      $ 2072 "Vial_liq_pick_3" "breakAfter"
      movel(Vial_liq_pick_3_p, a=0.5, v=0.1)
      $ 2073 "Vial_liq_pick_4" "breakAfter"
      movel(Vial_liq_pick_4_p, a=0.5, v=0.1)
      # begin: URCap Program Node
      #   Source: Robotiq_Grippers, 3.17.0.105337, Robotiq Inc.
      #   Type: Gripper
      $ 2074 "Gripper Close (1)"
      if not(gripper_connected[0]):
        popup("Gripper 1 must be connected to run this program.", "No connection", False, True, True)
      end
      if not(rq_is_gripper_activated("1")):
        popup("Gripper 1 is not activated. Go to Installation tab > Gripper to activate it and run the program again.", "Not activated", False, True, True)
      end
      rq_set_pos_spd_for(255, 82, 71, "1")
      rq_wait_pos_spe_for_request(255, 82, 71, "1")
      rq_go_to("1")
      rq_wait("1")
      # end: URCap Program Node
      $ 2075 "Wait: 1.0"
      sleep(1.0)
      $ 2076 "Set GRP_3F_Open=On"
      set_standard_digital_out(5, True)
      $ 2077 "Wait: 0.5"
      sleep(0.5)
      $ 2078 "Vial_liq_abov_2" "breakAfter"
      movel(Vial_liq_abov_2_p, a=0.3, v=0.05, r=0.05)
      $ 2079 "MoveL"
      $ 2080 "Liquid_midway_1" "breakAfter"
      movel(Liquid_midway_1_p, a=0.5, v=0.1)
      $ 2081 "Loop 3 times"
      Loop_1 = 0
      while (Loop_1 < 3):
        $ 2082 "shake_3" "breakAfter"
        movel(shake_3_p, a=2.0, v=0.5)
        $ 2083 "shake_4" "breakAfter"
        movel(shake_4_p, a=2.0, v=0.5)
        Loop_1 = Loop_1 + 1
      end
      $ 2084 "drop_above_3" "breakAfter"
      movel(drop_above_3_p, a=0.5, v=0.1)
      $ 2085 "drop_above_4" "breakAfter"
      movel(drop_above_4_p, a=0.5, v=0.1)
      $ 2086 "liq_tran_3" "breakAfter"
      movel(liq_tran_3_p, a=0.5, v=0.05, r=0.008)
      $ 2087 "Wait: 1.0"
      sleep(1.0)
      $ 2088 "drop_above_5" "breakAfter"
      movel(drop_above_5_p, a=0.5, v=0.1)
      $ 2089 "Waypoint_92" "breakAfter"
      movel(Waypoint_92_p, a=0.5, v=0.1)
      $ 2090 "liq_tran_4" "breakAfter"
      movel(liq_tran_4_p, a=0.5, v=0.05)
      $ 2091 "Wait: 1.0"
      sleep(1.0)
      $ 2092 "drop_above_6" "breakAfter"
      movel(drop_above_6_p, a=0.5, v=0.1)
      $ 2093 "drop_above_7" "breakAfter"
      movel(drop_above_7_p, a=0.5, v=0.1)
      $ 2094 "Liquid_midway_2" "breakAfter"
      movel(Liquid_midway_2_p, a=0.5, v=0.1)
      $ 2095 "MoveL"
      $ 2096 "Vial_drop_abo_1" "breakAfter"
      movel(Vial_drop_abo_1_p, a=0.5, v=0.1)
      $ 2097 "Vial_liq_drop_1" "breakAfter"
      movel(Vial_liq_drop_1_p, a=0.5, v=0.1)
      # begin: URCap Program Node
      #   Source: Robotiq_Grippers, 3.17.0.105337, Robotiq Inc.
      #   Type: Gripper
      $ 2098 "Gripper Open (1)"
      if not(gripper_connected[0]):
        popup("Gripper 1 must be connected to run this program.", "No connection", False, True, True)
      end
      if not(rq_is_gripper_activated("1")):
        popup("Gripper 1 is not activated. Go to Installation tab > Gripper to activate it and run the program again.", "Not activated", False, True, True)
      end
      rq_set_pos_spd_for(0, 82, 71, "1")
      rq_wait_pos_spe_for_request(0, 82, 71, "1")
      rq_go_to("1")
      rq_wait("1")
      # end: URCap Program Node
      $ 2099 "Vial_drop_abo_2" "breakAfter"
      movel(Vial_drop_abo_2_p, a=0.5, v=0.1)
    elif (34 == switch_1):
      $ 2100 "Case 34"
      $ 2101 "Task≔'Dosing'"
      global Task="Dosing"
      $ 2102 "tilt_to_home()"
      tilt_to_home()
      $ 2103 "Powder dosing all"
      $ 2104 "tilt_angle_sent≔0.0"
      global tilt_angle_sent=0.0
      $ 2105 "send_target_info()"
      send_target_info()
      $ 2107 "prev_spat≔''"
      global prev_spat=""
      $ 2108 "spatula≔''"
      global spatula=""
      $ 2109 "scoop_status≔'normal'"
      global scoop_status="normal"
      $ 2110 "send_powder_info()"
      send_powder_info()
      $ 2111 "Set AO[0]=0.0"
      set_standard_analog_out(0, 0.0)
      $ 2112 "Wait: 0.2"
      sleep(0.2)
      $ 2113 "reach pots decapping pose"
      # begin: URCap Program Node
      #   Source: SensoPart VISOR Robotic, 2.0.6, SensoPart Industriesensorik GmbH
      #   Type: VISOR Robotic App
      $ 2119 "VISOR Easy Pick"
      def visorFuncEasyPick_5caf8b():
        # begin: URCap Program Node
        #   Source: SensoPart VISOR Robotic, 2.0.6, SensoPart Industriesensorik GmbH
        #   Type: Easy Pick Setup
        $ 2120 "# 1 Setup" "noBreak"
        local easyPickVisorId = 1
        local easyPickArmMounted = True
        local easyPickSetJob = True
        local easyPickJobName = "Weight_scale"
        local easyPickAtImgAcq = False
        local easyPickImgAcqPose = Trigger
        # end: URCap Program Node
        # begin: URCap Program Node
        #   Source: SensoPart VISOR Robotic, 2.0.6, SensoPart Industriesensorik GmbH
        #   Type: Process
        $ 2121 "Process" "noBreak"
        local easyPickObjTaken = False
        local easyPickTrigger = False
        local easyPickPoseIdx = 0
        local easyPickPose = p[0,0,0,0,0,0]
        def easyPickFuncTrigger(visorId, setJob, jobName, arm):
        if (setJob):
          visor_changeJob(visorId, jobName, 6000)
        end
        if (arm):
          visor_trigger(visorId, 6000, "arm")
        else:
          visor_trigger(visorId, 6000)
        end
        global easyPickParts_4=visor_partsFound(visorId)
        visor_easyPickUpdate(visorId, "parts", visor_partsFound(visorId))
        return visor_getPose3d(visorId, 0)
      end
      while (not easyPickObjTaken):
        easyPickTrigger = (easyPickCount_4 >= visor_partsFound(easyPickVisorId)) or (easyPickCount_4 > 9) or (not visor_easyPickCheckIdent("a98771", easyPickVisorId))
        if (easyPickTrigger):
          easyPickCount_4 = 0
        end
        easyPickPoseIdx = easyPickCount_4
        easyPickPose = visor_getPose3d(easyPickVisorId, easyPickPoseIdx)
        visor_easyPickUpdate(easyPickVisorId, "counter", easyPickPoseIdx)
        # begin: URCap Program Node
        #   Source: SensoPart VISOR Robotic, 2.0.6, SensoPart Industriesensorik GmbH
        #   Type: Image Acquisition Pose
        $ 2122 "Image Acquisition Pose" "noBreak"
        if (easyPickTrigger):
          if (not easyPickAtImgAcq):
            movej(pose_trans(easyPickImgAcqPose,p[0.0000,0.0000,-0.0000,0.0000,0.0000,0.0000]),a=1.3963,v=1.0472,t=0.000000,r=0.000000)
            easyPickAtImgAcq = True
          end
          easyPickPose = easyPickFuncTrigger(easyPickVisorId, easyPickSetJob, easyPickJobName, easyPickArmMounted)
        end
        # end: URCap Program Node
        # begin: URCap Program Node
        #   Source: SensoPart VISOR Robotic, 2.0.6, SensoPart Industriesensorik GmbH
        #   Type: Object Detected
        $ 2123 "Object Detected" "noBreak"
        if (visor_partsFound(easyPickVisorId) > 0):
          $ 2124 "Open Gripper" "noBreak"
          $ 2125 "weight_value≔get_weight()" "noBreak"
          global weight_value=get_weight()
          $ 2126 "Wait: 0.5" "noBreak"
          sleep(0.5)
          $ 2127 "diff≔target_weight-weight_value" "noBreak"
          global diff=target_weight-weight_value
          $ 2128 "compute_level_percent(W_now, weight_value)" "noBreak"
          compute_level_percent(W_now, weight_value)
          $ 2129 "send_level_info()" "noBreak"
          send_level_info()
          $ 2130 "spatula≔select_spatula(Flowability, level, diff, bulk_density, mouth_d)" "noBreak"
          global spatula=select_spatula(Flowability, level, diff, bulk_density, mouth_d)
          $ 2131 "Wait: 0.2" "noBreak"
          sleep(0.2)
          $ 2132 "send_spatula_info()" "noBreak"
          send_spatula_info()
          $ 2133 "Pick spatula" "noBreak"
          $ 2134 "If spatula ≟ 'spatula_L'" "noBreak"
          if (spatula  ==  "spatula_L"):
            $ 2135 "MoveJ" "noBreak"
            $ 2136 "Spatula_otw" "noBreak"
            movej(get_inverse_kin(Spatula_otw_p, qnear=Spatula_otw_q), a=1.3962634015954636, v=1.0471975511965976)
            $ 2137 "pick_spat_L_abv" "noBreak"
            movej(get_inverse_kin(pick_spat_L_abv_p, qnear=pick_spat_L_abv_q), a=1.3962634015954636, v=1.0471975511965976)
            $ 2138 "MoveL" "noBreak"
            $ 2139 "spat_L_pick" "noBreak"
            movel(spat_L_pick_p, a=1.2, v=0.25)
            # begin: URCap Program Node
            #   Source: Robotiq_Grippers, 3.17.0.105337, Robotiq Inc.
            #   Type: Gripper
            $ 2140 "Gripper Close (1)" "noBreak"
            if not(gripper_connected[0]):
              popup("Gripper 1 must be connected to run this program.", "No connection", False, True, True)
            end
            if not(rq_is_gripper_activated("1")):
              popup("Gripper 1 is not activated. Go to Installation tab > Gripper to activate it and run the program again.", "Not activated", False, True, True)
            end
            rq_set_pos_spd_for(255, 0, 77, "1")
            rq_wait_pos_spe_for_request(255, 0, 77, "1")
            rq_go_to("1")
            rq_wait("1")
            # end: URCap Program Node
            $ 2141 "spat_L_lift" "noBreak"
            movel(spat_L_lift_p, a=1.2, v=0.25, r=0.01)
            $ 2142 "spat_L_side" "noBreak"
            movel(spat_L_side_p, a=1.2, v=0.25, r=0.01)
            $ 2143 "spat_L_up" "noBreak"
            movel(spat_L_up_p, a=1.2, v=0.25, r=0.05)
            $ 2144 "MoveJ" "noBreak"
            $ 2145 "Spatula_otw" "noBreak"
            movej(get_inverse_kin(Spatula_otw_p, qnear=Spatula_otw_q), a=1.3962634015954636, v=1.0471975511965976)
          else:
            $ 2146 "ElseIf spatula ≟'spatula_M'" "noBreak"
            if (spatula  == "spatula_M"):
              $ 2147 "MoveJ" "noBreak"
              $ 2148 "Spatula_otw" "noBreak"
              movej(get_inverse_kin(Spatula_otw_p, qnear=Spatula_otw_q), a=1.3962634015954636, v=1.0471975511965976)
              $ 2149 "spat_M_up" "noBreak"
              movej(get_inverse_kin(spat_M_up_p, qnear=spat_M_up_q), a=1.3962634015954636, v=1.0471975511965976, r=0.05)
              $ 2150 "MoveL" "noBreak"
              $ 2151 "spat_M_pick" "noBreak"
              movel(spat_M_pick_p, a=1.2, v=0.25)
              # begin: URCap Program Node
              #   Source: Robotiq_Grippers, 3.17.0.105337, Robotiq Inc.
              #   Type: Gripper
              $ 2152 "Gripper Close (1)" "noBreak"
              if not(gripper_connected[0]):
                popup("Gripper 1 must be connected to run this program.", "No connection", False, True, True)
              end
              if not(rq_is_gripper_activated("1")):
                popup("Gripper 1 is not activated. Go to Installation tab > Gripper to activate it and run the program again.", "Not activated", False, True, True)
              end
              rq_set_pos_spd_for(255, 0, 77, "1")
              rq_wait_pos_spe_for_request(255, 0, 77, "1")
              rq_go_to("1")
              rq_wait("1")
              # end: URCap Program Node
              $ 2153 "spat_M_up" "noBreak"
              movel(spat_M_up_p, a=1.2, v=0.25, r=0.05)
              $ 2154 "Spatula_otw" "noBreak"
              movel(Spatula_otw_p, a=1.2, v=0.25)
              $ 2155 "switch_spat_M≔ False " "noBreak"
              global switch_spat_M=  False
            else:
              $ 2156 "ElseIf spatula≟'spatula_S'" "noBreak"
              if (spatula == "spatula_S"):
                $ 2157 "MoveJ" "noBreak"
                $ 2158 "Spatula_otw" "noBreak"
                movej(get_inverse_kin(Spatula_otw_p, qnear=Spatula_otw_q), a=1.3962634015954636, v=1.0471975511965976)
                $ 2159 "spat_S_Up_7" "noBreak"
                movej(get_inverse_kin(spat_S_Up_7_p, qnear=spat_S_Up_7_q), a=1.3962634015954636, v=1.0471975511965976, r=0.05)
                $ 2160 "MoveL" "noBreak"
                $ 2161 "spat_S_Pick_4" "noBreak"
                movel(spat_S_Pick_4_p, a=1.2, v=0.25)
                # begin: URCap Program Node
                #   Source: Robotiq_Grippers, 3.17.0.105337, Robotiq Inc.
                #   Type: Gripper
                $ 2162 "Gripper Close (1)" "noBreak"
                if not(gripper_connected[0]):
                  popup("Gripper 1 must be connected to run this program.", "No connection", False, True, True)
                end
                if not(rq_is_gripper_activated("1")):
                  popup("Gripper 1 is not activated. Go to Installation tab > Gripper to activate it and run the program again.", "Not activated", False, True, True)
                end
                rq_set_pos_spd_for(255, 0, 77, "1")
                rq_wait_pos_spe_for_request(255, 0, 77, "1")
                rq_go_to("1")
                rq_wait("1")
                # end: URCap Program Node
                $ 2163 "spat_S_Up_8" "noBreak"
                movel(spat_S_Up_8_p, a=1.2, v=0.25, r=0.05)
                $ 2164 "Spatula_otw" "noBreak"
                movel(Spatula_otw_p, a=1.2, v=0.25)
                $ 2165 "switch_spat_S≔ False " "noBreak"
                global switch_spat_S=  False
              else:
                $ 2166 "ElseIf spatula≟'spatula_flat_M'" "noBreak"
                if (spatula == "spatula_flat_M"):
                  $ 2167 "MoveJ" "noBreak"
                  $ 2168 "Spatula_otw" "noBreak"
                  movej(get_inverse_kin(Spatula_otw_p, qnear=Spatula_otw_q), a=1.3962634015954636, v=1.0471975511965976)
                  $ 2169 "spat_flatM_up" "noBreak"
                  movej(get_inverse_kin(spat_flatM_up_p, qnear=spat_flatM_up_q), a=1.3962634015954636, v=1.0471975511965976, r=0.05)
                  $ 2170 "MoveL" "noBreak"
                  $ 2171 "spat_flatM_pick" "noBreak"
                  movel(spat_flatM_pick_p, a=1.2, v=0.25)
                  # begin: URCap Program Node
                  #   Source: Robotiq_Grippers, 3.17.0.105337, Robotiq Inc.
                  #   Type: Gripper
                  $ 2172 "Gripper Close (1)" "noBreak"
                  if not(gripper_connected[0]):
                    popup("Gripper 1 must be connected to run this program.", "No connection", False, True, True)
                  end
                  if not(rq_is_gripper_activated("1")):
                    popup("Gripper 1 is not activated. Go to Installation tab > Gripper to activate it and run the program again.", "Not activated", False, True, True)
                  end
                  rq_set_pos_spd_for(255, 0, 77, "1")
                  rq_wait_pos_spe_for_request(255, 0, 77, "1")
                  rq_go_to("1")
                  rq_wait("1")
                  # end: URCap Program Node
                  $ 2173 "spat_flatM_up" "noBreak"
                  movel(spat_flatM_up_p, a=1.2, v=0.25, r=0.05)
                  $ 2174 "Spatula_otw" "noBreak"
                  movel(Spatula_otw_p, a=1.2, v=0.25)
                  $ 2175 "switch_spat_F_M≔ False " "noBreak"
                  global switch_spat_F_M=  False
                else:
                  $ 2176 "ElseIf spatula≟'spatula_flat_S'" "noBreak"
                  if (spatula == "spatula_flat_S"):
                    $ 2177 "MoveJ" "noBreak"
                    $ 2178 "Spatula_otw" "noBreak"
                    movej(get_inverse_kin(Spatula_otw_p, qnear=Spatula_otw_q), a=1.3962634015954636, v=1.0471975511965976)
                    $ 2179 "spat_flatS_up" "noBreak"
                    movej(get_inverse_kin(spat_flatS_up_p, qnear=spat_flatS_up_q), a=1.3962634015954636, v=1.0471975511965976, r=0.05)
                    $ 2180 "MoveL" "noBreak"
                    $ 2181 "spat_flatS_pick" "noBreak"
                    movel(spat_flatS_pick_p, a=1.2, v=0.25)
                    # begin: URCap Program Node
                    #   Source: Robotiq_Grippers, 3.17.0.105337, Robotiq Inc.
                    #   Type: Gripper
                    $ 2182 "Gripper Close (1)" "noBreak"
                    if not(gripper_connected[0]):
                      popup("Gripper 1 must be connected to run this program.", "No connection", False, True, True)
                    end
                    if not(rq_is_gripper_activated("1")):
                      popup("Gripper 1 is not activated. Go to Installation tab > Gripper to activate it and run the program again.", "Not activated", False, True, True)
                    end
                    rq_set_pos_spd_for(255, 0, 77, "1")
                    rq_wait_pos_spe_for_request(255, 0, 77, "1")
                    rq_go_to("1")
                    rq_wait("1")
                    # end: URCap Program Node
                    $ 2183 "spat_flatS_up" "noBreak"
                    movel(spat_flatS_up_p, a=1.2, v=0.25, r=0.05)
                    $ 2184 "Spatula_otw" "noBreak"
                    movel(Spatula_otw_p, a=1.2, v=0.25)
                    $ 2185 "switch_spat_F_S≔ False " "noBreak"
                    global switch_spat_F_S=  False
                  end
                end
              end
            end
          end
          $ 2186 "Action_Info≔'Scooping'" "noBreak"
          global Action_Info="Scooping"
          $ 2187 "auto_tilt_and_scoop(W_now, target_weight, weight_value)" "noBreak"
          auto_tilt_and_scoop(W_now, target_weight, weight_value)
          $ 2188 "Action_Info≔'Dosing'" "noBreak"
          global Action_Info="Dosing"
          # begin: URCap Program Node
          #   Source: SensoPart VISOR Robotic, 2.0.6, SensoPart Industriesensorik GmbH
          #   Type: Approach Pose
          $ 2189 "Approach Pose" "noBreak"
          movej(pose_trans(easyPickPose,p[0.0000,0.0000,-0.0000,0.0000,0.0000,0.0000]),a=0.2618,v=0.1745,t=0.000000,r=0.000000)
          # end: URCap Program Node
          # begin: URCap Program Node
          #   Source: SensoPart VISOR Robotic, 2.0.6, SensoPart Industriesensorik GmbH
          #   Type: Target Pose
          $ 2190 "Target Pose" "noBreak"
          movel(pose_trans(easyPickPose,p[0.0000,0.0000,-0.0000,0.0000,0.0000,0.0000]),a=0.0500,v=0.0200,t=0.000000,r=0.000000)
          # end: URCap Program Node
          $ 2191 "Close Gripper" "noBreak"
          $ 2192 "current_p≔get_actual_tcp_pose()" "noBreak"
          global current_p= get_actual_tcp_pose ()
          $ 2193 "dispense_pos≔pose_trans(current_p,p[0,0,0,0,-deg2rad(spatula_ry),0])" "noBreak"
          global dispense_pos=pose_trans(current_p,p[0,0,0,0,-deg2rad(spatula_ry),0])
          $ 2195 "Loop weight_value≤target_weight " "noBreak"
          thread Thread_while_2195():
            while (True):
              $ 2196 "MoveL" "noBreak"
              $ 2197 "dispense_pos" "noBreak"
              movel(dispense_pos, a=0.2, v=0.1)
              $ 2198 "log_weight()" "noBreak"
              log_weight()
              $ 2200 "CCW_full_Rotate()" "noBreak"
              CCW_full_Rotate()
              $ 2201 "Start_thread≔ True " "noBreak"
              global Start_thread=  True
              $ 2202 "vib_thread≔ True " "noBreak"
              global vib_thread=  True
              $ 2203 "Wait: 0.5" "noBreak"
              sleep(0.5)
              $ 2204 "If diff ≥(target_g*1.2)" "noBreak"
              if (diff  >= (target_g*1.2)):
                $ 2205 "tilt_pose≔pose_trans(get_actual_tcp_pose(), p[0, 0, 0, 0, 0, 2.0])" "noBreak"
                global tilt_pose=pose_trans(get_actual_tcp_pose(), p[0, 0, 0, 0, 0, 2.0])
                $ 2206 "movel(tilt_pose, a=0.5, v=0.5, r=0.00001)" "noBreak"
                movel(tilt_pose, a=0.5, v=0.5, r=0.00001)
              else:
                $ 2207 "Else" "noBreak"
                $ 2208 "Loop weight_value≤(target_weight-0.00) and tilt_angle≥(-1.999) and tilt_angle≤0.5" "noBreak"
                thread Thread_while_2208():
                  while (True):
                    $ 2209 "current_error≔target_weight-weight_value" "noBreak"
                    global current_error=target_weight-weight_value
                    $ 2210 "Integral_error≔Integral_error+current_error*dt" "noBreak"
                    global Integral_error=Integral_error+current_error*dt
                    $ 2211 "derivative≔(current_error-previous_error)/dt" "noBreak"
                    global derivative=(current_error-previous_error)/dt
                    $ 2212 "tilt_increment≔(kp*current_error)+(ki*Integral_error)+(kd*derivative)" "noBreak"
                    global tilt_increment=(kp*current_error)+(ki*Integral_error)+(kd*derivative)
                    $ 2213 "current_pose≔get_actual_tcp_pose()" "noBreak"
                    global current_pose= get_actual_tcp_pose ()
                    $ 2214 "tilt_angle≔current_pose[5]" "noBreak"
                    global tilt_angle=current_pose[5]
                    $ 2215 "tilt_pose≔pose_trans(current_pose, p[0, 0, 0, 0, 0, tilt_increment])" "noBreak"
                    global tilt_pose=pose_trans(current_pose, p[0, 0, 0, 0, 0, tilt_increment])
                    $ 2216 "movel(tilt_pose, a=0.1, v=0.1, r=0.00001)" "noBreak"
                    movel(tilt_pose, a=0.1, v=0.1, r=0.00001)
                    $ 2217 "previous_error≔current_error" "noBreak"
                    global previous_error=current_error
                  end
                end
                if (weight_value <= (target_weight-0.00)  and  tilt_angle >= (-1.999)  and  tilt_angle <= 0.5):
                  global thread_handler_2208=run Thread_while_2208()
                  while (weight_value <= (target_weight-0.00)  and  tilt_angle >= (-1.999)  and  tilt_angle <= 0.5):
                    sync()
                  end
                  kill thread_handler_2208
                end
              end
              $ 2218 "weight_value≔get_weight()" "noBreak"
              global weight_value=get_weight()
              $ 2220 "tilt_angle≔-1" "noBreak"
              global tilt_angle=-1
              $ 2221 "Wait: 0.5" "noBreak"
              sleep(0.5)
              $ 2222 "Start_thread≔ False " "noBreak"
              global Start_thread=  False
              $ 2223 "vib_thread≔ False " "noBreak"
              global vib_thread=  False
              $ 2225 "dispense_pos" "noBreak"
              movel(dispense_pos, a=1.2, v=0.25)
              $ 2226 "compute_level_percent(W_now, weight_value)" "noBreak"
              compute_level_percent(W_now, weight_value)
              $ 2227 "prev_spat≔spatula" "noBreak"
              global prev_spat=spatula
              $ 2228 "Wait: 0.2" "noBreak"
              sleep(0.2)
              $ 2229 "spatula≔select_spatula(Flowability, level, diff, bulk_density, mouth_d)" "noBreak"
              global spatula=select_spatula(Flowability, level, diff, bulk_density, mouth_d)
              $ 2230 "Wait: 1.0" "noBreak"
              sleep(1.0)
              $ 2231 "send_level_info()" "noBreak"
              send_level_info()
              $ 2232 "send_spatula_info()" "noBreak"
              send_spatula_info()
              $ 2233 "Integral_error≔0" "noBreak"
              global Integral_error=0
              $ 2234 "current_error≔0" "noBreak"
              global current_error=0
              $ 2235 "previous_error≔0" "noBreak"
              global previous_error=0
              $ 2236 "Set AO[0]=0.0" "noBreak"
              set_standard_analog_out(0, 0.0)
              $ 2237 "Wait: 0.5" "noBreak"
              sleep(0.5)
              $ 2238 "swtich spatula" "noBreak"
              $ 2239 "If spatula ≟ 'spatula_M' and switch_spat_M≟ True " "noBreak"
              if (spatula  ==  "spatula_M"  and  switch_spat_M ==   True  ):
                $ 2240 "MoveJ" "noBreak"
                $ 2241 "Spatula_otw" "noBreak"
                movej(get_inverse_kin(Spatula_otw_p, qnear=Spatula_otw_q), a=1.3962634015954636, v=1.0471975511965976)
                $ 2242 "spat_L_up" "noBreak"
                movej(get_inverse_kin(spat_L_up_p, qnear=spat_L_up_q), a=1.3962634015954636, v=1.0471975511965976)
                $ 2243 "MoveL" "noBreak"
                $ 2244 "spat_L_side" "noBreak"
                movel(spat_L_side_p, a=1.2, v=0.25)
                $ 2245 "spat_L_lift" "noBreak"
                movel(spat_L_lift_p, a=1.2, v=0.25)
                $ 2246 "spat_L_pick" "noBreak"
                movel(spat_L_pick_p, a=0.2, v=0.1)
                # begin: URCap Program Node
                #   Source: Robotiq_Grippers, 3.17.0.105337, Robotiq Inc.
                #   Type: Gripper
                $ 2247 "Gripper Open (1)" "noBreak"
                if not(gripper_connected[0]):
                  popup("Gripper 1 must be connected to run this program.", "No connection", False, True, True)
                end
                if not(rq_is_gripper_activated("1")):
                  popup("Gripper 1 is not activated. Go to Installation tab > Gripper to activate it and run the program again.", "Not activated", False, True, True)
                end
                rq_set_pos_spd_for(0, 255, 77, "1")
                rq_wait_pos_spe_for_request(0, 255, 77, "1")
                rq_go_to("1")
                rq_wait("1")
                # end: URCap Program Node
                $ 2248 "spat_M_pick" "noBreak"
                movel(spat_M_pick_p, a=1.2, v=0.25)
                # begin: URCap Program Node
                #   Source: Robotiq_Grippers, 3.17.0.105337, Robotiq Inc.
                #   Type: Gripper
                $ 2249 "Gripper Close (1)" "noBreak"
                if not(gripper_connected[0]):
                  popup("Gripper 1 must be connected to run this program.", "No connection", False, True, True)
                end
                if not(rq_is_gripper_activated("1")):
                  popup("Gripper 1 is not activated. Go to Installation tab > Gripper to activate it and run the program again.", "Not activated", False, True, True)
                end
                rq_set_pos_spd_for(255, 0, 77, "1")
                rq_wait_pos_spe_for_request(255, 0, 77, "1")
                rq_go_to("1")
                rq_wait("1")
                # end: URCap Program Node
                $ 2250 "spat_M_up" "noBreak"
                movel(spat_M_up_p, a=1.2, v=0.25)
                $ 2251 "Spatula_otw" "noBreak"
                movel(Spatula_otw_p, a=1.2, v=0.25)
                $ 2252 "switch_spat_M≔ False " "noBreak"
                global switch_spat_M=  False
                $ 2253 "correction_reset()" "noBreak"
                correction_reset()
              else:
                $ 2254 "ElseIf spatula ≟ 'spatula_S' and switch_spat_S ≟ True and prev_spat≟'spatula_M'" "noBreak"
                if (spatula  ==  "spatula_S" and switch_spat_S  ==   True  and prev_spat == "spatula_M"):
                  $ 2255 "MoveL" "noBreak"
                  $ 2256 "Spatula_otw" "noBreak"
                  movel(Spatula_otw_p, a=1.2, v=0.25)
                  $ 2257 "spat_M_up" "noBreak"
                  movel(spat_M_up_p, a=1.2, v=0.25)
                  $ 2258 "spat_M_pick" "noBreak"
                  movel(spat_M_pick_p, a=0.2, v=0.1)
                  # begin: URCap Program Node
                  #   Source: Robotiq_Grippers, 3.17.0.105337, Robotiq Inc.
                  #   Type: Gripper
                  $ 2259 "Gripper Open (1)" "noBreak"
                  if not(gripper_connected[0]):
                    popup("Gripper 1 must be connected to run this program.", "No connection", False, True, True)
                  end
                  if not(rq_is_gripper_activated("1")):
                    popup("Gripper 1 is not activated. Go to Installation tab > Gripper to activate it and run the program again.", "Not activated", False, True, True)
                  end
                  rq_set_pos_spd_for(0, 255, 77, "1")
                  rq_wait_pos_spe_for_request(0, 255, 77, "1")
                  rq_go_to("1")
                  rq_wait("1")
                  # end: URCap Program Node
                  $ 2260 "spat_S_pick" "noBreak"
                  movel(spat_S_pick_p, a=1.2, v=0.25)
                  # begin: URCap Program Node
                  #   Source: Robotiq_Grippers, 3.17.0.105337, Robotiq Inc.
                  #   Type: Gripper
                  $ 2261 "Gripper Close (1)" "noBreak"
                  if not(gripper_connected[0]):
                    popup("Gripper 1 must be connected to run this program.", "No connection", False, True, True)
                  end
                  if not(rq_is_gripper_activated("1")):
                    popup("Gripper 1 is not activated. Go to Installation tab > Gripper to activate it and run the program again.", "Not activated", False, True, True)
                  end
                  rq_set_pos_spd_for(255, 0, 77, "1")
                  rq_wait_pos_spe_for_request(255, 0, 77, "1")
                  rq_go_to("1")
                  rq_wait("1")
                  # end: URCap Program Node
                  $ 2262 "spat_S_up" "noBreak"
                  movel(spat_S_up_p, a=1.2, v=0.25)
                  $ 2263 "Spatula_otw" "noBreak"
                  movel(Spatula_otw_p, a=1.2, v=0.25)
                  $ 2264 "switch_spat_S≔ False " "noBreak"
                  global switch_spat_S=  False
                  $ 2265 "correction_reset()" "noBreak"
                  correction_reset()
                else:
                  $ 2266 "ElseIf spatula≟'spatula_S' and switch_spat_S≟ True  and prev_spat≟'spatula_L'" "noBreak"
                  if (spatula == "spatula_S" and switch_spat_S ==   True    and  prev_spat == "spatula_L"):
                    $ 2267 "MoveJ" "noBreak"
                    $ 2268 "Spatula_otw" "noBreak"
                    movej(get_inverse_kin(Spatula_otw_p, qnear=Spatula_otw_q), a=1.3962634015954636, v=1.0471975511965976)
                    $ 2269 "spat_L_up" "noBreak"
                    movej(get_inverse_kin(spat_L_up_p, qnear=spat_L_up_q), a=1.3962634015954636, v=1.0471975511965976)
                    $ 2270 "MoveL" "noBreak"
                    $ 2271 "spat_L_side" "noBreak"
                    movel(spat_L_side_p, a=1.2, v=0.25)
                    $ 2272 "spat_L_lift" "noBreak"
                    movel(spat_L_lift_p, a=1.2, v=0.25)
                    $ 2273 "spat_L_pick" "noBreak"
                    movel(spat_L_pick_p, a=0.2, v=0.1)
                    # begin: URCap Program Node
                    #   Source: Robotiq_Grippers, 3.17.0.105337, Robotiq Inc.
                    #   Type: Gripper
                    $ 2274 "Gripper Open (1)" "noBreak"
                    if not(gripper_connected[0]):
                      popup("Gripper 1 must be connected to run this program.", "No connection", False, True, True)
                    end
                    if not(rq_is_gripper_activated("1")):
                      popup("Gripper 1 is not activated. Go to Installation tab > Gripper to activate it and run the program again.", "Not activated", False, True, True)
                    end
                    rq_set_pos_spd_for(0, 255, 77, "1")
                    rq_wait_pos_spe_for_request(0, 255, 77, "1")
                    rq_go_to("1")
                    rq_wait("1")
                    # end: URCap Program Node
                    $ 2275 "spat_S_pick" "noBreak"
                    movel(spat_S_pick_p, a=1.2, v=0.25)
                    # begin: URCap Program Node
                    #   Source: Robotiq_Grippers, 3.17.0.105337, Robotiq Inc.
                    #   Type: Gripper
                    $ 2276 "Gripper Close (1)" "noBreak"
                    if not(gripper_connected[0]):
                      popup("Gripper 1 must be connected to run this program.", "No connection", False, True, True)
                    end
                    if not(rq_is_gripper_activated("1")):
                      popup("Gripper 1 is not activated. Go to Installation tab > Gripper to activate it and run the program again.", "Not activated", False, True, True)
                    end
                    rq_set_pos_spd_for(255, 0, 77, "1")
                    rq_wait_pos_spe_for_request(255, 0, 77, "1")
                    rq_go_to("1")
                    rq_wait("1")
                    # end: URCap Program Node
                    $ 2277 "spat_S_up" "noBreak"
                    movel(spat_S_up_p, a=1.2, v=0.25)
                    $ 2278 "Spatula_otw" "noBreak"
                    movel(Spatula_otw_p, a=1.2, v=0.25)
                    $ 2279 "switch_spat_S≔ False " "noBreak"
                    global switch_spat_S=  False
                    $ 2280 "correction_reset()" "noBreak"
                    correction_reset()
                  else:
                    $ 2281 "ElseIf spatula≟'spatula_flat_S'  and switch_spat_F_S ≟ True " "noBreak"
                    if (spatula == "spatula_flat_S"   and  switch_spat_F_S  ==   True  ):
                      $ 2282 "MoveL" "noBreak"
                      $ 2283 "Spatula_otw" "noBreak"
                      movel(Spatula_otw_p, a=1.2, v=0.25)
                      $ 2284 "spat_flatM_up" "noBreak"
                      movel(spat_flatM_up_p, a=1.2, v=0.25)
                      $ 2285 "spat_flatM_pick" "noBreak"
                      movel(spat_flatM_pick_p, a=0.2, v=0.1)
                      # begin: URCap Program Node
                      #   Source: Robotiq_Grippers, 3.17.0.105337, Robotiq Inc.
                      #   Type: Gripper
                      $ 2286 "Gripper Open (1)" "noBreak"
                      if not(gripper_connected[0]):
                        popup("Gripper 1 must be connected to run this program.", "No connection", False, True, True)
                      end
                      if not(rq_is_gripper_activated("1")):
                        popup("Gripper 1 is not activated. Go to Installation tab > Gripper to activate it and run the program again.", "Not activated", False, True, True)
                      end
                      rq_set_pos_spd_for(0, 255, 74, "1")
                      rq_wait_pos_spe_for_request(0, 255, 74, "1")
                      rq_go_to("1")
                      rq_wait("1")
                      # end: URCap Program Node
                      $ 2287 "spat_flatS_pick" "noBreak"
                      movel(spat_flatS_pick_p, a=1.2, v=0.25)
                      # begin: URCap Program Node
                      #   Source: Robotiq_Grippers, 3.17.0.105337, Robotiq Inc.
                      #   Type: Gripper
                      $ 2288 "Gripper Close (1)" "noBreak"
                      if not(gripper_connected[0]):
                        popup("Gripper 1 must be connected to run this program.", "No connection", False, True, True)
                      end
                      if not(rq_is_gripper_activated("1")):
                        popup("Gripper 1 is not activated. Go to Installation tab > Gripper to activate it and run the program again.", "Not activated", False, True, True)
                      end
                      rq_set_pos_spd_for(255, 0, 77, "1")
                      rq_wait_pos_spe_for_request(255, 0, 77, "1")
                      rq_go_to("1")
                      rq_wait("1")
                      # end: URCap Program Node
                      $ 2289 "spat_flatS_up" "noBreak"
                      movel(spat_flatS_up_p, a=1.2, v=0.25)
                      $ 2290 "Spatula_otw" "noBreak"
                      movel(Spatula_otw_p, a=1.2, v=0.25)
                      $ 2291 "switch_spat_F_S≔ False " "noBreak"
                      global switch_spat_F_S=  False
                      $ 2292 "correction_reset()" "noBreak"
                      correction_reset()
                    end
                  end
                end
              end
              $ 2293 "tilt(level)" "noBreak"
              tilt(level)
              $ 2294 "Action_Info≔'Scooping'" "noBreak"
              global Action_Info="Scooping"
              $ 2295 "auto_tilt_and_scoop(W_now, target_weight, weight_value)" "noBreak"
              auto_tilt_and_scoop(W_now, target_weight, weight_value)
              $ 2296 "Action_Info≔'Dosing'" "noBreak"
              global Action_Info="Dosing"
            end
          end
          if (weight_value <= target_weight ):
            global thread_handler_2195=run Thread_while_2195()
            while (weight_value <= target_weight ):
              sync()
            end
            kill thread_handler_2195
          end
          $ 2297 "Start_thread≔ False " "noBreak"
          global Start_thread=  False
          $ 2298 "vib_thread≔ False " "noBreak"
          global vib_thread=  False
          # begin: URCap Program Node
          #   Source: SensoPart VISOR Robotic, 2.0.6, SensoPart Industriesensorik GmbH
          #   Type: Exit Pose
          $ 2299 "Exit Pose" "noBreak"
          movel(pose_trans(easyPickPose,p[0.0000,0.0000,-0.0000,0.0000,0.0000,0.0000]),a=0.5000,v=0.2500,t=0.000000,r=0.000000)
          # end: URCap Program Node
          easyPickObjTaken = True
        end
        # end: URCap Program Node
        # begin: URCap Program Node
        #   Source: SensoPart VISOR Robotic, 2.0.6, SensoPart Industriesensorik GmbH
        #   Type: No Object Detected
        $ 2300 "No Object Detected" "noBreak"
        if (visor_partsFound(easyPickVisorId) < 1):
          $ 2301 "Popup: No weigh scale detected" "noBreak"
          popup("No weigh scale detected", "Message", False, False, blocking=True)
          else:
        end
        # end: URCap Program Node
      end
      easyPickCount_4 = easyPickCount_4 + 1
      visor_easyPickUpdate(easyPickVisorId, "counter", easyPickCount_4)
      visor_easyPickSetIdent("a98771", easyPickVisorId)
      # end: URCap Program Node
    end
    visorFuncEasyPick_5caf8b()
    # end: URCap Program Node
    $ 2302 "MoveL"
    $ 2303 "dispense_pos" "breakAfter"
    movel(dispense_pos, a=0.2, v=0.1)
    $ 2304 "after_scoop()"
    after_scoop()
    $ 2305 "Place spatula back to the rack"
    $ 2306 "If spatula ≟ 'spatula_L'"
    if (spatula  ==  "spatula_L"):
      $ 2307 "MoveJ"
      $ 2308 "Spatula_otw" "breakAfter"
      movej(get_inverse_kin(Spatula_otw_p, qnear=Spatula_otw_q), a=1.3962634015954636, v=1.0471975511965976)
      $ 2309 "MoveL"
      $ 2310 "spat_L_up" "breakAfter"
      movel(spat_L_up_p, a=1.2, v=0.25, r=0.05)
      $ 2311 "spat_L_side" "breakAfter"
      movel(spat_L_side_p, a=1.2, v=0.25, r=0.01)
      $ 2312 "spat_L_lift" "breakAfter"
      movel(spat_L_lift_p, a=1.2, v=0.25, r=0.01)
      $ 2313 "spat_L_pick" "breakAfter"
      movel(spat_L_pick_p, a=0.2, v=0.1)
      # begin: URCap Program Node
      #   Source: Robotiq_Grippers, 3.17.0.105337, Robotiq Inc.
      #   Type: Gripper
      $ 2314 "Gripper Open (1)"
      if not(gripper_connected[0]):
        popup("Gripper 1 must be connected to run this program.", "No connection", False, True, True)
      end
      if not(rq_is_gripper_activated("1")):
        popup("Gripper 1 is not activated. Go to Installation tab > Gripper to activate it and run the program again.", "Not activated", False, True, True)
      end
      rq_set_pos_spd_for(0, 128, 128, "1")
      rq_wait_pos_spe_for_request(0, 128, 128, "1")
      rq_go_to("1")
      rq_wait("1")
      # end: URCap Program Node
      $ 2315 "MoveJ"
      $ 2316 "pick_spat_L_abv" "breakAfter"
      movej(get_inverse_kin(pick_spat_L_abv_p, qnear=pick_spat_L_abv_q), a=1.3962634015954636, v=1.0471975511965976)
      $ 2317 "Spatula_otw" "breakAfter"
      movej(get_inverse_kin(Spatula_otw_p, qnear=Spatula_otw_q), a=1.3962634015954636, v=1.0471975511965976)
    else:
      $ 2318 "ElseIf spatula ≟'spatula_M'"
      if (spatula  == "spatula_M"):
        $ 2319 "MoveJ"
        $ 2320 "Spatula_otw" "breakAfter"
        movej(get_inverse_kin(Spatula_otw_p, qnear=Spatula_otw_q), a=1.3962634015954636, v=1.0471975511965976)
        $ 2321 "spat_M_up" "breakAfter"
        movej(get_inverse_kin(spat_M_up_p, qnear=spat_M_up_q), a=1.3962634015954636, v=1.0471975511965976, r=0.05)
        $ 2322 "MoveL"
        $ 2323 "spat_M_pick" "breakAfter"
        movel(spat_M_pick_p, a=0.2, v=0.1)
        # begin: URCap Program Node
        #   Source: Robotiq_Grippers, 3.17.0.105337, Robotiq Inc.
        #   Type: Gripper
        $ 2324 "Gripper Open (1)"
        if not(gripper_connected[0]):
          popup("Gripper 1 must be connected to run this program.", "No connection", False, True, True)
        end
        if not(rq_is_gripper_activated("1")):
          popup("Gripper 1 is not activated. Go to Installation tab > Gripper to activate it and run the program again.", "Not activated", False, True, True)
        end
        rq_set_pos_spd_for(0, 128, 128, "1")
        rq_wait_pos_spe_for_request(0, 128, 128, "1")
        rq_go_to("1")
        rq_wait("1")
        # end: URCap Program Node
        $ 2325 "spat_M_up" "breakAfter"
        movel(spat_M_up_p, a=1.2, v=0.25, r=0.05)
        $ 2326 "Spatula_otw" "breakAfter"
        movel(Spatula_otw_p, a=1.2, v=0.25)
        $ 2327 "switch_spat_M≔ False "
        global switch_spat_M=  False
      else:
        $ 2328 "ElseIf spatula≟'spatula_S'"
        if (spatula == "spatula_S"):
          $ 2329 "MoveJ"
          $ 2330 "Spatula_otw" "breakAfter"
          movej(get_inverse_kin(Spatula_otw_p, qnear=Spatula_otw_q), a=1.3962634015954636, v=1.0471975511965976)
          $ 2331 "spat_S_Up_7" "breakAfter"
          movej(get_inverse_kin(spat_S_Up_7_p, qnear=spat_S_Up_7_q), a=1.3962634015954636, v=1.0471975511965976, r=0.05)
          $ 2332 "MoveL"
          $ 2333 "spat_S_Pick_4" "breakAfter"
          movel(spat_S_Pick_4_p, a=0.2, v=0.1)
          # begin: URCap Program Node
          #   Source: Robotiq_Grippers, 3.17.0.105337, Robotiq Inc.
          #   Type: Gripper
          $ 2334 "Gripper Open (1)"
          if not(gripper_connected[0]):
            popup("Gripper 1 must be connected to run this program.", "No connection", False, True, True)
          end
          if not(rq_is_gripper_activated("1")):
            popup("Gripper 1 is not activated. Go to Installation tab > Gripper to activate it and run the program again.", "Not activated", False, True, True)
          end
          rq_set_pos_spd_for(0, 255, 51, "1")
          rq_wait_pos_spe_for_request(0, 255, 51, "1")
          rq_go_to("1")
          rq_wait("1")
          # end: URCap Program Node
          $ 2335 "spat_S_Up_8" "breakAfter"
          movel(spat_S_Up_8_p, a=1.2, v=0.25, r=0.05)
          $ 2336 "Spatula_otw" "breakAfter"
          movel(Spatula_otw_p, a=1.2, v=0.25)
          $ 2337 "switch_spat_S≔ False "
          global switch_spat_S=  False
        else:
          $ 2338 "ElseIf spatula≟'spatula_flat_M'"
          if (spatula == "spatula_flat_M"):
            $ 2339 "MoveJ"
            $ 2340 "Spatula_otw" "breakAfter"
            movej(get_inverse_kin(Spatula_otw_p, qnear=Spatula_otw_q), a=1.3962634015954636, v=1.0471975511965976)
            $ 2341 "spat_flatM_up" "breakAfter"
            movej(get_inverse_kin(spat_flatM_up_p, qnear=spat_flatM_up_q), a=1.3962634015954636, v=1.0471975511965976, r=0.05)
            $ 2342 "MoveL"
            $ 2343 "spat_flatM_pick" "breakAfter"
            movel(spat_flatM_pick_p, a=0.2, v=0.1)
            # begin: URCap Program Node
            #   Source: Robotiq_Grippers, 3.17.0.105337, Robotiq Inc.
            #   Type: Gripper
            $ 2344 "Gripper Open (1)"
            if not(gripper_connected[0]):
              popup("Gripper 1 must be connected to run this program.", "No connection", False, True, True)
            end
            if not(rq_is_gripper_activated("1")):
              popup("Gripper 1 is not activated. Go to Installation tab > Gripper to activate it and run the program again.", "Not activated", False, True, True)
            end
            rq_set_pos_spd_for(0, 128, 128, "1")
            rq_wait_pos_spe_for_request(0, 128, 128, "1")
            rq_go_to("1")
            rq_wait("1")
            # end: URCap Program Node
            $ 2345 "spat_flatM_up" "breakAfter"
            movel(spat_flatM_up_p, a=1.2, v=0.25, r=0.05)
            $ 2346 "Spatula_otw" "breakAfter"
            movel(Spatula_otw_p, a=1.2, v=0.25)
            $ 2347 "switch_spat_F_M≔ False "
            global switch_spat_F_M=  False
          else:
            $ 2348 "ElseIf spatula≟'spatula_flat_S'"
            if (spatula == "spatula_flat_S"):
              $ 2349 "MoveJ"
              $ 2350 "Spatula_otw" "breakAfter"
              movej(get_inverse_kin(Spatula_otw_p, qnear=Spatula_otw_q), a=1.3962634015954636, v=1.0471975511965976)
              $ 2351 "spat_flatS_up" "breakAfter"
              movej(get_inverse_kin(spat_flatS_up_p, qnear=spat_flatS_up_q), a=1.3962634015954636, v=1.0471975511965976, r=0.05)
              $ 2352 "MoveL"
              $ 2353 "spat_flatS_pick" "breakAfter"
              movel(spat_flatS_pick_p, a=0.2, v=0.1)
              # begin: URCap Program Node
              #   Source: Robotiq_Grippers, 3.17.0.105337, Robotiq Inc.
              #   Type: Gripper
              $ 2354 "Gripper Open (1)"
              if not(gripper_connected[0]):
                popup("Gripper 1 must be connected to run this program.", "No connection", False, True, True)
              end
              if not(rq_is_gripper_activated("1")):
                popup("Gripper 1 is not activated. Go to Installation tab > Gripper to activate it and run the program again.", "Not activated", False, True, True)
              end
              rq_set_pos_spd_for(0, 128, 128, "1")
              rq_wait_pos_spe_for_request(0, 128, 128, "1")
              rq_go_to("1")
              rq_wait("1")
              # end: URCap Program Node
              $ 2355 "spat_flatS_up" "breakAfter"
              movel(spat_flatS_up_p, a=1.2, v=0.25, r=0.05)
              $ 2356 "Spatula_otw" "breakAfter"
              movel(Spatula_otw_p, a=1.2, v=0.25)
              $ 2357 "switch_spat_F_S≔ False "
              global switch_spat_F_S=  False
            end
          end
        end
      end
    end
    $ 2358 "switch_spat_M≔ True "
    global switch_spat_M=  True
    $ 2359 "switch_spat_S≔ True "
    global switch_spat_S=  True
    $ 2360 "switch_spat_F_M≔ True "
    global switch_spat_F_M=  True
    $ 2361 "switch_spat_F_S≔ True "
    global switch_spat_F_S=  True
    $ 2362 "correction_reset()"
    correction_reset()
  elif (38 == switch_1):
    $ 2558 "Case 38"
    $ 2559 "Decap Powder container"
    $ 2560 "MoveJ"
    $ 2562 "Waypoint_7" "breakAfter"
    movej(get_inverse_kin(Waypoint_7_p, qnear=Waypoint_7_q), a=1.3962634015954636, v=1.0471975511965976, r=0.05)
    $ 2563 "MoveL"
    $ 2565 "Waypoint_8" "breakAfter"
    movel(Waypoint_8_p, a=1.2, v=0.25)
    $ 2566 "MoveL"
    $ 2567 "Decapp_above_3" "breakAfter"
    movel(Decapp_above_3_p, a=1.2, v=0.25)
    $ 2568 "Set GRP_3F_Open=On"
    set_standard_digital_out(5, True)
    $ 2569 "Wait: 0.5"
    sleep(0.5)
    $ 2570 "Decapp_place_3" "breakAfter"
    movel(Decapp_place_3_p, a=0.3, v=0.05)
    $ 2571 "Set GRP_3F_Open=Off"
    set_standard_digital_out(5, False)
    $ 2572 "Wait: 0.5"
    sleep(0.5)
    # begin: URCap Program Node
    #   Source: Robotiq_Grippers, 3.17.0.105337, Robotiq Inc.
    #   Type: Gripper
    $ 2573 "Gripper Open (1)"
    if not(gripper_connected[0]):
      popup("Gripper 1 must be connected to run this program.", "No connection", False, True, True)
    end
    if not(rq_is_gripper_activated("1")):
      popup("Gripper 1 is not activated. Go to Installation tab > Gripper to activate it and run the program again.", "Not activated", False, True, True)
    end
    rq_set_pos_spd_for(0, 77, 77, "1")
    rq_wait_pos_spe_for_request(0, 77, 77, "1")
    rq_go_to("1")
    rq_wait("1")
    # end: URCap Program Node
    $ 2574 "MoveL"
    $ 2575 "Decapp_above_4" "breakAfter"
    movel(Decapp_above_4_p, a=1.2, v=0.25)
    $ 2576 "Waypoint_78" "breakAfter"
    movel(Waypoint_78_p, a=1.2, v=0.25, r=0.05)
    $ 2577 "Home (Safe)"
    movej([-1.2302089344500047, -1.2969853503591224, -1.875639182904262, -1.539621866126728, 1.5731943360401213, -2.80099559440227], a=1.3962634015954636, v=1.0471975511965976)
  elif (39 == switch_1):
    $ 2578 "Case 39"
    $ 2579 "Powder container Pick"
    $ 2580 "Direct Pick"
    $ 2581 "Set"
    set_tcp(p[0.0,0.0,0.15052000000000001,3.1415,0.0,0.0])
    $ 2582 "read_db_data()"
    read_db_data()
    # begin: URCap Program Node
    #   Source: SensoPart VISOR Robotic, 2.0.6, SensoPart Industriesensorik GmbH
    #   Type: VISOR ChangeJob
    $ 2583 "# 1 VISOR ChangeJob"
    visor_changeJob(1, "Aztec_no_dot_pick", 6000)
    # end: URCap Program Node
    # begin: URCap Program Node
    #   Source: SensoPart VISOR Robotic, 2.0.6, SensoPart Industriesensorik GmbH
    #   Type: VISOR Terminal
    $ 2584 "# 1 VISOR Terminal"
    visor_terminal(1, "TRX00", 3000)
    # end: URCap Program Node
    $ 2585 "table_pick_TCP≔visor_getPose3d(1, 0)"
    global table_pick_TCP= visor_getPose3d (1, 0)
    # begin: URCap Program Node
    #   Source: Robotiq_Grippers, 3.17.0.105337, Robotiq Inc.
    #   Type: Gripper
    $ 2586 "Gripper Open (1)"
    if not(gripper_connected[0]):
      popup("Gripper 1 must be connected to run this program.", "No connection", False, True, True)
    end
    if not(rq_is_gripper_activated("1")):
      popup("Gripper 1 is not activated. Go to Installation tab > Gripper to activate it and run the program again.", "Not activated", False, True, True)
    end
    rq_set_pos_spd_for(0, 77, 77, "1")
    rq_wait_pos_spe_for_request(0, 77, 77, "1")
    rq_go_to("1")
    rq_wait("1")
    # end: URCap Program Node
    $ 2587 "MoveJ"
    $ 2589 "Waypoint_10" "breakAfter"
    movej(get_inverse_kin(Waypoint_10_p, qnear=Waypoint_10_q), a=1.3962634015954636, v=1.0471975511965976, r=0.05)
    $ 2590 "Waypoint_9" "breakAfter"
    movej(get_inverse_kin(Waypoint_9_p, qnear=Waypoint_9_q), a=1.3962634015954636, v=1.0471975511965976, r=0.05)
    $ 2591 "MoveJ"
    $ 2593 "table_prepick≔pose_trans(table_pick_TCP,p[0,0,cent_edge/2,0,0,0])"
    global table_prepick=pose_trans(table_pick_TCP,p[0,0,cent_edge/2,0,0,0])
    $ 2594 "table_prepick" "breakAfter"
    movej(table_prepick, a=0.8726646259971648, v=0.6981317007977318)
    $ 2595 "table_safe_pick≔pose_trans(table_prepick, p[0,pick_2_base-H_c,cent_edge/2,0,0,0])"
    global table_safe_pick= pose_trans (table_prepick, p[0,pick_2_base-H_c,cent_edge/2,0,0,0])
    $ 2596 "table_safe_pick" "breakAfter"
    movej(table_safe_pick, a=0.8726646259971648, v=0.6981317007977318, r=0.05)
    $ 2597 "table_pick≔pose_trans(table_prepick, p[0,pick_2_base - d_cc,0,0,0,0])"
    global table_pick= pose_trans (table_prepick, p[0,pick_2_base - d_cc,0,0,0,0])
    $ 2598 "table_pick" "breakAfter"
    movej(table_pick, a=0.8726646259971648, v=0.6981317007977318)
    # begin: URCap Program Node
    #   Source: Robotiq_Grippers, 3.17.0.105337, Robotiq Inc.
    #   Type: Gripper
    $ 2599 "Gripper Close (1)"
    if not(gripper_connected[0]):
      popup("Gripper 1 must be connected to run this program.", "No connection", False, True, True)
    end
    if not(rq_is_gripper_activated("1")):
      popup("Gripper 1 is not activated. Go to Installation tab > Gripper to activate it and run the program again.", "Not activated", False, True, True)
    end
    rq_set_pos_spd_for(255, 77, 51, "1")
    rq_wait_pos_spe_for_request(255, 77, 51, "1")
    rq_go_to("1")
    rq_wait("1")
    # end: URCap Program Node
    $ 2600 "table_prepick" "breakAfter"
    movej(table_prepick, a=0.8726646259971648, v=0.6981317007977318)
    $ 2601 "Picking≔ True "
    global Picking=  True
    $ 2631 "powder_position≔'Position2'"
    global powder_position="Position2"
    $ 2632 "MoveJ"
    $ 2633 "Powder_wayp1" "breakAfter"
    movej(get_inverse_kin(Powder_wayp1_p, qnear=Powder_wayp1_q), a=1.3962634015954636, v=1.0471975511965976, r=0.05)
    $ 2634 "MoveL"
    $ 2635 "Waypoint_2" "breakAfter"
    movel(Waypoint_2_p, a=1.2, v=0.25)
    $ 2636 "Set"
    set_tcp(p[0.0,0.0,0.161,3.1415,0.0,0.0])
    $ 2637 "If powder_position ≟ 'Position1'"
    if (powder_position  ==  "Position1"):
      $ 2638 "MoveJ"
      $ 2639 "Postions_otw" "breakAfter"
      movej(get_inverse_kin(Postions_otw_p, qnear=Postions_otw_q), a=1.3962634015954636, v=1.0471975511965976, r=0.01)
      $ 2640 "MoveL"
      $ 2641 "Cont_A_TCP" "breakAfter"
      movel(Cont_A_TCP, a=0.5, v=0.2)
      $ 2642 "cont_A_prepick≔pose_trans(Cont_A_TCP, p[0,0,cent_edge/2,0,0,0])"
      global cont_A_prepick= pose_trans (Cont_A_TCP, p[0,0,cent_edge/2,0,0,0])
      $ 2643 "cont_A_prepick" "breakAfter"
      movel(cont_A_prepick, a=0.3, v=0.05)
      $ 2644 "cont_A_pick≔pose_trans(cont_A_prepick, p[0,pick_2_base-d_cc,0,0,0,0])"
      global cont_A_pick= pose_trans (cont_A_prepick, p[0,pick_2_base-d_cc,0,0,0,0])
      $ 2645 "cont_A_pick" "breakAfter"
      movel(cont_A_pick, a=0.2, v=0.1)
      # begin: URCap Program Node
      #   Source: Robotiq_Grippers, 3.17.0.105337, Robotiq Inc.
      #   Type: Gripper
      $ 2646 "Gripper Open (1)"
      if not(gripper_connected[0]):
        popup("Gripper 1 must be connected to run this program.", "No connection", False, True, True)
      end
      if not(rq_is_gripper_activated("1")):
        popup("Gripper 1 is not activated. Go to Installation tab > Gripper to activate it and run the program again.", "Not activated", False, True, True)
      end
      rq_set_pos_spd_for(0, 77, 26, "1")
      rq_wait_pos_spe_for_request(0, 77, 26, "1")
      rq_go_to("1")
      rq_wait("1")
      # end: URCap Program Node
      $ 2647 "cont_A_otw" "breakAfter"
      movel(cont_A_otw_p, a=0.5, v=0.2)
      $ 2648 "cont_A_prepick" "breakAfter"
      movel(cont_A_prepick, a=0.5, v=0.2)
      $ 2649 "Postions_otw" "breakAfter"
      movel(Postions_otw_p, a=0.5, v=0.2, r=0.01)
      $ 2651 "Home (Safe)"
      movej([-1.2302089344500047, -1.2969853503591224, -1.875639182904262, -1.539621866126728, 1.5731943360401213, -2.80099559440227], a=1.3962634015954636, v=1.0471975511965976)
    else:
      $ 2653 "ElseIf powder_position≟'Position2'"
      if (powder_position == "Position2"):
        $ 2654 "MoveJ"
        $ 2655 "Postions_otw" "breakAfter"
        movej(get_inverse_kin(Postions_otw_p, qnear=Postions_otw_q), a=1.3962634015954636, v=1.0471975511965976, r=0.01)
        $ 2656 "MoveL"
        $ 2659 "cont_B_prepick≔pose_trans(Cont_B_TCP, p[0,0,cent_edge/2,0,0,0])"
        global cont_B_prepick= pose_trans (Cont_B_TCP, p[0,0,cent_edge/2,0,0,0])
        $ 2660 "cont_B_prepick" "breakAfter"
        movel(cont_B_prepick, a=1.2, v=0.25)
        $ 2661 "cont_B_pick≔pose_trans(cont_B_prepick, p[0,pick_2_base-d_cc,0,0,0,0])"
        global cont_B_pick= pose_trans (cont_B_prepick, p[0,pick_2_base-d_cc,0,0,0,0])
        $ 2662 "cont_B_pick" "breakAfter"
        global move_thread_flag_2662=0
        thread move_thread_2662():
          enter_critical
          move_thread_flag_2662 = 1
          movel(cont_B_pick, a=0.2, v=0.1)
          move_thread_flag_2662 = 2
          exit_critical
        end
        move_thread_flag_2662 = 0
        move_thread_han_2662 = run move_thread_2662()
        while (True):
          local targetTcpDirection=get_target_tcp_speed()
          local stepsToRetract=tool_contact(direction=targetTcpDirection, force_threshold=8.000000)
          if (stepsToRetract > 0):
            kill move_thread_han_2662
            stopl(3.0)
            local backTrackMovement=get_actual_joint_positions_history(stepsToRetract)
            local contactPose=get_forward_kin(backTrackMovement)
            local posDir=[targetTcpDirection[0],targetTcpDirection[1],targetTcpDirection[2]]
            local retractTo=contactPose
            if (norm(posDir) > 1e-6):
              local normalizedPosDir=normalize(posDir)
              local additionalRetraction=p[normalizedPosDir[0] * 0.0, normalizedPosDir[1] * 0.0, normalizedPosDir[2] * 0.0, 0, 0, 0]
              retractTo = pose_sub(contactPose, additionalRetraction)
            end
            movel(retractTo, a=3.0, v=0.1)
            $ 2663 "Until (tool_contact_detection)"
            $ 2664 "saved_place_pos≔get_actual_tcp_pose()"
            global saved_place_pos= get_actual_tcp_pose ()
            break
          end
          sleep(1.0E-10)
          if (move_thread_flag_2662 > 1):
            join move_thread_han_2662
            break
          end
          sync()
        end
        # begin: URCap Program Node
        #   Source: Robotiq_Grippers, 3.17.0.105337, Robotiq Inc.
        #   Type: Gripper
        $ 2665 "Gripper Open (1)"
        if not(gripper_connected[0]):
          popup("Gripper 1 must be connected to run this program.", "No connection", False, True, True)
        end
        if not(rq_is_gripper_activated("1")):
          popup("Gripper 1 is not activated. Go to Installation tab > Gripper to activate it and run the program again.", "Not activated", False, True, True)
        end
        rq_set_pos_spd_for(0, 77, 26, "1")
        rq_wait_pos_spe_for_request(0, 77, 26, "1")
        rq_go_to("1")
        rq_wait("1")
        # end: URCap Program Node
        $ 2666 "cont_B_otw" "breakAfter"
        movel(cont_B_otw_p, a=1.2, v=0.25)
        $ 2668 "cont_B_safe" "breakAfter"
        movel(cont_B_safe_p, a=1.2, v=0.25)
        $ 2669 "Postions_otw" "breakAfter"
        movel(Postions_otw_p, a=1.2, v=0.25)
        $ 2670 "Home (Safe)"
        movej([-1.2302089344500047, -1.2969853503591224, -1.875639182904262, -1.539621866126728, 1.5731943360401213, -2.80099559440227], a=1.3962634015954636, v=1.0471975511965976)
      else:
        $ 2672 "ElseIf powder_position≟'Position3'"
        if (powder_position == "Position3"):
          $ 2673 "MoveJ"
          $ 2674 "Postions_otw" "breakAfter"
          movej(get_inverse_kin(Postions_otw_p, qnear=Postions_otw_q), a=1.3962634015954636, v=1.0471975511965976, r=0.01)
          $ 2681 "MoveL"
          $ 2682 "Cont_C_TCP" "breakAfter"
          movel(Cont_C_TCP, a=1.2, v=0.25, r=0.01)
          $ 2683 "cont_C_prepick≔pose_trans(Cont_C_TCP, p[0,0,cent_edge/2,0,0,0])"
          global cont_C_prepick= pose_trans (Cont_C_TCP, p[0,0,cent_edge/2,0,0,0])
          $ 2684 "cont_C_prepick" "breakAfter"
          movel(cont_C_prepick, a=0.3, v=0.05)
          $ 2685 "cont_C_pick≔pose_trans(cont_C_prepick, p[0,pick_2_base-d_cc,0,0,0,0])"
          global cont_C_pick= pose_trans (cont_C_prepick, p[0,pick_2_base-d_cc,0,0,0,0])
          $ 2686 "cont_C_pick" "breakAfter"
          movel(cont_C_pick, a=0.2, v=0.1)
          # begin: URCap Program Node
          #   Source: Robotiq_Grippers, 3.17.0.105337, Robotiq Inc.
          #   Type: Gripper
          $ 2687 "Gripper Open (1)"
          if not(gripper_connected[0]):
            popup("Gripper 1 must be connected to run this program.", "No connection", False, True, True)
          end
          if not(rq_is_gripper_activated("1")):
            popup("Gripper 1 is not activated. Go to Installation tab > Gripper to activate it and run the program again.", "Not activated", False, True, True)
          end
          rq_set_pos_spd_for(0, 77, 26, "1")
          rq_wait_pos_spe_for_request(0, 77, 26, "1")
          rq_go_to("1")
          rq_wait("1")
          # end: URCap Program Node
          $ 2688 "cont_C_otw" "breakAfter"
          movel(cont_C_otw_p, a=1.2, v=0.25)
          $ 2689 "cont_C_prepick" "breakAfter"
          movel(cont_C_prepick, a=1.2, v=0.25, r=0.01)
          $ 2690 "Postions_otw" "breakAfter"
          movel(Postions_otw_p, a=1.2, v=0.25)
          $ 2691 "Home (Safe)"
          movej([-1.2302089344500047, -1.2969853503591224, -1.875639182904262, -1.539621866126728, 1.5731943360401213, -2.80099559440227], a=1.3962634015954636, v=1.0471975511965976)
        end
      end
    end
    $ 2693 "Home (Safe)"
    movej([-1.2302089344500047, -1.2969853503591224, -1.875639182904262, -1.539621866126728, 1.5731943360401213, -2.80099559440227], a=1.3962634015954636, v=1.0471975511965976)
  elif (41 == switch_1):
    $ 2802 "Case 41"
    $ 2803 "Task≔'Decapping_Dosing'"
    global Task="Decapping_Dosing"
    $ 2804 "tilt_to_home()"
    tilt_to_home()
    $ 2805 "Weigh, Place & decap container"
    $ 2806 "Set"
    set_tcp(p[0.0,0.0,0.15052000000000001,3.1415,0.0,0.0])
    # begin: URCap Program Node
    #   Source: SensoPart VISOR Robotic, 2.0.6, SensoPart Industriesensorik GmbH
    #   Type: VISOR Robotic App
    $ 2807 "VISOR Easy Pick"
    def visorFuncEasyPick_44508e():
      # begin: URCap Program Node
      #   Source: SensoPart VISOR Robotic, 2.0.6, SensoPart Industriesensorik GmbH
      #   Type: Easy Pick Setup
      $ 2808 "# 1 Setup" "noBreak"
      local easyPickVisorId = 1
      local easyPickArmMounted = True
      local easyPickSetJob = True
      local easyPickJobName = "PoTS"
      local easyPickAtImgAcq = False
      local easyPickImgAcqPose = FRM_PoTS
      # end: URCap Program Node
      # begin: URCap Program Node
      #   Source: SensoPart VISOR Robotic, 2.0.6, SensoPart Industriesensorik GmbH
      #   Type: Process
      $ 2809 "Process" "noBreak"
      local easyPickObjTaken = False
      local easyPickTrigger = False
      local easyPickPoseIdx = 0
      local easyPickPose = p[0,0,0,0,0,0]
      def easyPickFuncTrigger(visorId, setJob, jobName, arm):
      if (setJob):
        visor_changeJob(visorId, jobName, 6000)
      end
      if (arm):
        visor_trigger(visorId, 6000, "arm")
      else:
        visor_trigger(visorId, 6000)
      end
      global easyPickParts_7=visor_partsFound(visorId)
      visor_easyPickUpdate(visorId, "parts", visor_partsFound(visorId))
      return visor_getPose3d(visorId, 0)
    end
    while (not easyPickObjTaken):
      easyPickTrigger = (easyPickCount_7 >= visor_partsFound(easyPickVisorId)) or (easyPickCount_7 > 9) or (not visor_easyPickCheckIdent("f0f0e4", easyPickVisorId))
      if (easyPickTrigger):
        easyPickCount_7 = 0
      end
      easyPickPoseIdx = easyPickCount_7
      easyPickPose = visor_getPose3d(easyPickVisorId, easyPickPoseIdx)
      visor_easyPickUpdate(easyPickVisorId, "counter", easyPickPoseIdx)
      # begin: URCap Program Node
      #   Source: SensoPart VISOR Robotic, 2.0.6, SensoPart Industriesensorik GmbH
      #   Type: Image Acquisition Pose
      $ 2810 "Image Acquisition Pose" "noBreak"
      if (easyPickTrigger):
        if (not easyPickAtImgAcq):
          movej(pose_trans(easyPickImgAcqPose,p[0.0000,0.0000,-0.0000,0.0000,0.0000,0.0000]),a=1.3963,v=1.0472,t=0.000000,r=0.000000)
          easyPickAtImgAcq = True
        end
        easyPickPose = easyPickFuncTrigger(easyPickVisorId, easyPickSetJob, easyPickJobName, easyPickArmMounted)
      end
      # end: URCap Program Node
      # begin: URCap Program Node
      #   Source: SensoPart VISOR Robotic, 2.0.6, SensoPart Industriesensorik GmbH
      #   Type: Object Detected
      $ 2811 "Object Detected" "noBreak"
      if (visor_partsFound(easyPickVisorId) > 0):
        $ 2812 "Open Gripper" "noBreak"
        # begin: URCap Program Node
        #   Source: Robotiq_Grippers, 3.17.0.105337, Robotiq Inc.
        #   Type: Gripper
        $ 2813 "Gripper Open (1)" "noBreak"
        if not(gripper_connected[0]):
          popup("Gripper 1 must be connected to run this program.", "No connection", False, True, True)
        end
        if not(rq_is_gripper_activated("1")):
          popup("Gripper 1 is not activated. Go to Installation tab > Gripper to activate it and run the program again.", "Not activated", False, True, True)
        end
        rq_set_pos_spd_for(0, 77, 77, "1")
        rq_wait_pos_spe_for_request(0, 77, 77, "1")
        rq_go_to("1")
        rq_wait("1")
        # end: URCap Program Node
        $ 2814 "Set" "noBreak"
        set_tcp(p[0.0,0.0,0.161,3.1415,0.0,0.0])
        $ 2815 "Wait: 0.2" "noBreak"
        sleep(0.2)
        $ 2816 "Place on second weigh scale" "noBreak"
        $ 2817 "MoveJ" "noBreak"
        $ 2818 "Waypoint_1" "noBreak"
        movej(get_inverse_kin(Waypoint_1_p, qnear=Waypoint_1_q), a=1.3962634015954636, v=1.0471975511965976, r=0.1)
        $ 2819 "Waypoint_5" "noBreak"
        movej(get_inverse_kin(Waypoint_5_p, qnear=Waypoint_5_q), a=1.3962634015954636, v=1.0471975511965976)
        $ 2821 "If Picking≟ True " "noBreak"
        if (Picking ==   True  ):
          $ 2822 "Pick from saved pose" "noBreak"
          $ 2823 "MoveL" "noBreak"
          $ 2824 "cont_B_safe" "noBreak"
          movel(cont_B_safe_p, a=0.2, v=0.1)
          $ 2825 "saved_place_pos" "noBreak"
          movel(saved_place_pos, a=1.2, v=0.25)
          # begin: URCap Program Node
          #   Source: Robotiq_Grippers, 3.17.0.105337, Robotiq Inc.
          #   Type: Gripper
          $ 2826 "Gripper Close (1)" "noBreak"
          if not(gripper_connected[0]):
            popup("Gripper 1 must be connected to run this program.", "No connection", False, True, True)
          end
          if not(rq_is_gripper_activated("1")):
            popup("Gripper 1 is not activated. Go to Installation tab > Gripper to activate it and run the program again.", "Not activated", False, True, True)
          end
          rq_set_pos_spd_for(255, 77, 26, "1")
          rq_wait_pos_spe_for_request(255, 77, 26, "1")
          rq_go_to("1")
          rq_wait("1")
          # end: URCap Program Node
          $ 2827 "cont_B_safe" "noBreak"
          movel(cont_B_safe_p, a=1.2, v=0.25)
          $ 2828 "Postions_otw" "noBreak"
          movel(Postions_otw_p, a=1.2, v=0.25)
        else:
          $ 2831 "Else" "noBreak"
          $ 2832 "read_db_data()" "noBreak"
          read_db_data()
          $ 2833 "Pick from B" "noBreak"
          $ 2834 "MoveL" "noBreak"
          $ 2836 "cont_B_safe" "noBreak"
          movel(cont_B_safe_p, a=1.2, v=0.25)
          $ 2837 "cont_B_prepick≔pose_trans(Cont_B_TCP, p[0,0,cent_edge/2,0,0,0])" "noBreak"
          global cont_B_prepick= pose_trans (Cont_B_TCP, p[0,0,cent_edge/2,0,0,0])
          $ 2838 "cont_B_otw" "noBreak"
          movel(cont_B_otw_p, a=1.2, v=0.25)
          $ 2840 "cont_B_pick≔pose_trans(cont_B_prepick, p[0,pick_2_base-d_cc,0,0,0,0])" "noBreak"
          global cont_B_pick= pose_trans (cont_B_prepick, p[0,pick_2_base-d_cc,0,0,0,0])
          $ 2841 "cont_B_pick" "noBreak"
          movel(cont_B_pick, a=0.2, v=0.1)
          # begin: URCap Program Node
          #   Source: Robotiq_Grippers, 3.17.0.105337, Robotiq Inc.
          #   Type: Gripper
          $ 2842 "Gripper Close (1)" "noBreak"
          if not(gripper_connected[0]):
            popup("Gripper 1 must be connected to run this program.", "No connection", False, True, True)
          end
          if not(rq_is_gripper_activated("1")):
            popup("Gripper 1 is not activated. Go to Installation tab > Gripper to activate it and run the program again.", "Not activated", False, True, True)
          end
          rq_set_pos_spd_for(255, 77, 51, "1")
          rq_wait_pos_spe_for_request(255, 77, 51, "1")
          rq_go_to("1")
          rq_wait("1")
          # end: URCap Program Node
          $ 2843 "cont_B_prepick" "noBreak"
          movel(cont_B_prepick, a=1.2, v=0.25, r=0.01)
          $ 2844 "Postions_otw" "noBreak"
          movel(Postions_otw_p, a=1.2, v=0.25)
        end
        $ 2861 "Set" "noBreak"
        set_tcp(p[0.0,0.0,0.15052000000000001,3.1415,0.0,0.0])
        # begin: URCap Program Node
        #   Source: SensoPart VISOR Robotic, 2.0.6, SensoPart Industriesensorik GmbH
        #   Type: Approach Pose
        $ 2862 "Approach Pose" "noBreak"
        movej(pose_trans(easyPickPose,p[0.0000,0.0000,-0.0000,0.0000,0.0000,0.0000]),a=0.5236,v=0.4363,t=0.000000,r=0.000000)
        # end: URCap Program Node
        # begin: URCap Program Node
        #   Source: SensoPart VISOR Robotic, 2.0.6, SensoPart Industriesensorik GmbH
        #   Type: Target Pose
        $ 2863 "Target Pose" "noBreak"
        movel(pose_trans(easyPickPose,p[0.0000,0.0000,-0.0000,0.0000,0.0000,0.0000]),a=0.1000,v=0.0500,t=0.000000,r=0.000000)
        # end: URCap Program Node
        $ 2864 "Close Gripper" "noBreak"
        $ 2865 "container_place≔get_actual_tcp_pose()" "noBreak"
        global container_place= get_actual_tcp_pose ()
        $ 2866 "PoTS_place_abov≔pose_trans(container_place, p[0,0,cent_edge/2,0,0,0])" "noBreak"
        global PoTS_place_abov=pose_trans(container_place, p[0,0,cent_edge/2,0,0,0])
        $ 2867 "MoveL" "noBreak"
        $ 2868 "PoTS_place_abov" "noBreak"
        movel(PoTS_place_abov, a=0.5, v=0.05)
        $ 2870 "target_pose≔pose_trans(PoTS_place_abov, p[0,pick_2_base-d_cc,0,0,0,0])" "noBreak"
        global target_pose=pose_trans(PoTS_place_abov, p[0,pick_2_base-d_cc,0,0,0,0])
        $ 2871 "MoveL" "noBreak"
        $ 2872 "target_pose" "noBreak"
        movel(target_pose, a=0.3, v=0.05)
        # begin: URCap Program Node
        #   Source: Robotiq_Grippers, 3.17.0.105337, Robotiq Inc.
        #   Type: Gripper
        $ 2873 "Gripper Open (1)" "noBreak"
        if not(gripper_connected[0]):
          popup("Gripper 1 must be connected to run this program.", "No connection", False, True, True)
        end
        if not(rq_is_gripper_activated("1")):
          popup("Gripper 1 is not activated. Go to Installation tab > Gripper to activate it and run the program again.", "Not activated", False, True, True)
        end
        rq_set_pos_spd_for(0, 77, 77, "1")
        rq_wait_pos_spe_for_request(0, 77, 77, "1")
        rq_go_to("1")
        rq_wait("1")
        # end: URCap Program Node
        # begin: URCap Program Node
        #   Source: SensoPart VISOR Robotic, 2.0.6, SensoPart Industriesensorik GmbH
        #   Type: Exit Pose
        $ 2874 "Exit Pose" "noBreak"
        movel(pose_trans(easyPickPose,p[0.0000,0.0000,0.1000,0.0000,0.0000,0.0000]),a=0.5000,v=0.2500,t=0.000000,r=0.000000)
        # end: URCap Program Node
        easyPickObjTaken = True
      end
      # end: URCap Program Node
      # begin: URCap Program Node
      #   Source: SensoPart VISOR Robotic, 2.0.6, SensoPart Industriesensorik GmbH
      #   Type: No Object Detected
      $ 2875 "No Object Detected" "noBreak"
      if (visor_partsFound(easyPickVisorId) < 1):
        $ 2876 "Popup: No POTS detected" "noBreak"
        popup("No POTS detected", "Message", False, False, blocking=True)
        else:
      end
      # end: URCap Program Node
    end
    easyPickCount_7 = easyPickCount_7 + 1
    visor_easyPickUpdate(easyPickVisorId, "counter", easyPickCount_7)
    visor_easyPickSetIdent("f0f0e4", easyPickVisorId)
    # end: URCap Program Node
  end
  visorFuncEasyPick_44508e()
  # end: URCap Program Node
  $ 2911 "MoveJ"
  $ 2912 "place_2_home" "breakAfter"
  movej(get_inverse_kin(place_2_home_p, qnear=place_2_home_q), a=1.3962634015954636, v=1.0471975511965976)
  $ 2913 "Picking≔ False "
  global Picking=  False
  elif (42 == switch_1):
    $ 2914 "Case 42"
  elif (43 == switch_1):
    $ 3676 "Case 43"
  elif (44 == switch_1):
    $ 3929 "Case 44"
  elif (45 == switch_1):
    $ 3993 "Case 45"
  elif (46 == switch_1):
    $ 4030 "Case 46"
  elif (47 == switch_1):
    $ 4320 "Case 47"
  elif (48 == switch_1):
    $ 4375 "Case 48"
  elif (49 == switch_1):
    $ 4393 "Case 49"
  elif (50 == switch_1):
    $ 4411 "Case 50"
    $ 4412 "Emptying powder container"
    $ 4413 "tilt_to_home()"
    tilt_to_home()
    $ 4414 "scoop_status≔'emptying'"
    global scoop_status="emptying"
    $ 4415 "Dosing untill empty"
    $ 4416 "tilt_angle_sent≔0.0"
    global tilt_angle_sent=0.0
    $ 4417 "send_target_info()"
    send_target_info()
    $ 4418 "zero_scale()"
    zero_scale()
    $ 4419 "prev_spat≔''"
    global prev_spat=""
    $ 4420 "spatula≔''"
    global spatula=""
    $ 4421 "send_powder_info()"
    send_powder_info()
    $ 4422 "Set AO[0]=0.0"
    set_standard_analog_out(0, 0.0)
    $ 4423 "Wait: 0.2"
    sleep(0.2)
    $ 4424 "reach pots decapping pose"
    # begin: URCap Program Node
    #   Source: SensoPart VISOR Robotic, 2.0.6, SensoPart Industriesensorik GmbH
    #   Type: VISOR Robotic App
    $ 4430 "VISOR Easy Pick"
    def visorFuncEasyPick_45d1f0():
      # begin: URCap Program Node
      #   Source: SensoPart VISOR Robotic, 2.0.6, SensoPart Industriesensorik GmbH
      #   Type: Easy Pick Setup
      $ 4431 "# 1 Setup" "noBreak"
      local easyPickVisorId = 1
      local easyPickArmMounted = True
      local easyPickSetJob = True
      local easyPickJobName = "Weight_scale"
      local easyPickAtImgAcq = False
      local easyPickImgAcqPose = Trigger
      # end: URCap Program Node
      # begin: URCap Program Node
      #   Source: SensoPart VISOR Robotic, 2.0.6, SensoPart Industriesensorik GmbH
      #   Type: Process
      $ 4432 "Process" "noBreak"
      local easyPickObjTaken = False
      local easyPickTrigger = False
      local easyPickPoseIdx = 0
      local easyPickPose = p[0,0,0,0,0,0]
      def easyPickFuncTrigger(visorId, setJob, jobName, arm):
      if (setJob):
        visor_changeJob(visorId, jobName, 6000)
      end
      if (arm):
        visor_trigger(visorId, 6000, "arm")
      else:
        visor_trigger(visorId, 6000)
      end
      global easyPickParts_4=visor_partsFound(visorId)
      visor_easyPickUpdate(visorId, "parts", visor_partsFound(visorId))
      return visor_getPose3d(visorId, 0)
    end
    while (not easyPickObjTaken):
      easyPickTrigger = (easyPickCount_4 >= visor_partsFound(easyPickVisorId)) or (easyPickCount_4 > 9) or (not visor_easyPickCheckIdent("cf4c8f", easyPickVisorId))
      if (easyPickTrigger):
        easyPickCount_4 = 0
      end
      easyPickPoseIdx = easyPickCount_4
      easyPickPose = visor_getPose3d(easyPickVisorId, easyPickPoseIdx)
      visor_easyPickUpdate(easyPickVisorId, "counter", easyPickPoseIdx)
      # begin: URCap Program Node
      #   Source: SensoPart VISOR Robotic, 2.0.6, SensoPart Industriesensorik GmbH
      #   Type: Image Acquisition Pose
      $ 4433 "Image Acquisition Pose" "noBreak"
      if (easyPickTrigger):
        if (not easyPickAtImgAcq):
          movej(pose_trans(easyPickImgAcqPose,p[0.0000,0.0000,-0.0000,0.0000,0.0000,0.0000]),a=1.3963,v=1.0472,t=0.000000,r=0.000000)
          easyPickAtImgAcq = True
        end
        easyPickPose = easyPickFuncTrigger(easyPickVisorId, easyPickSetJob, easyPickJobName, easyPickArmMounted)
      end
      # end: URCap Program Node
      # begin: URCap Program Node
      #   Source: SensoPart VISOR Robotic, 2.0.6, SensoPart Industriesensorik GmbH
      #   Type: Object Detected
      $ 4434 "Object Detected" "noBreak"
      if (visor_partsFound(easyPickVisorId) > 0):
        $ 4435 "Open Gripper" "noBreak"
        $ 4436 "weight_value≔get_weight()" "noBreak"
        global weight_value=get_weight()
        $ 4437 "Wait: 1.0" "noBreak"
        sleep(1.0)
        $ 4438 "diff≔target_weight-weight_value" "noBreak"
        global diff=target_weight-weight_value
        $ 4439 "compute_level_percent(W_now, weight_value)" "noBreak"
        compute_level_percent(W_now, weight_value)
        $ 4440 "send_level_info()" "noBreak"
        send_level_info()
        $ 4441 "spatula≔select_spatula(Flowability, level, diff, bulk_density, mouth_d)" "noBreak"
        global spatula=select_spatula(Flowability, level, diff, bulk_density, mouth_d)
        $ 4442 "Wait: 0.2" "noBreak"
        sleep(0.2)
        $ 4443 "send_spatula_info()" "noBreak"
        send_spatula_info()
        $ 4444 "Pick spatula" "noBreak"
        $ 4445 "If spatula ≟ 'spatula_L'" "noBreak"
        if (spatula  ==  "spatula_L"):
          $ 4446 "MoveJ" "noBreak"
          $ 4447 "Spatula_otw" "noBreak"
          movej(get_inverse_kin(Spatula_otw_p, qnear=Spatula_otw_q), a=1.3962634015954636, v=1.0471975511965976)
          $ 4448 "pick_spat_L_abv" "noBreak"
          movej(get_inverse_kin(pick_spat_L_abv_p, qnear=pick_spat_L_abv_q), a=1.3962634015954636, v=1.0471975511965976)
          $ 4449 "MoveL" "noBreak"
          $ 4450 "spat_L_pick" "noBreak"
          movel(spat_L_pick_p, a=1.2, v=0.25)
          # begin: URCap Program Node
          #   Source: Robotiq_Grippers, 3.17.0.105337, Robotiq Inc.
          #   Type: Gripper
          $ 4451 "Gripper Close (1)" "noBreak"
          if not(gripper_connected[0]):
            popup("Gripper 1 must be connected to run this program.", "No connection", False, True, True)
          end
          if not(rq_is_gripper_activated("1")):
            popup("Gripper 1 is not activated. Go to Installation tab > Gripper to activate it and run the program again.", "Not activated", False, True, True)
          end
          rq_set_pos_spd_for(255, 0, 77, "1")
          rq_wait_pos_spe_for_request(255, 0, 77, "1")
          rq_go_to("1")
          rq_wait("1")
          # end: URCap Program Node
          $ 4452 "spat_L_lift" "noBreak"
          movel(spat_L_lift_p, a=1.2, v=0.25, r=0.01)
          $ 4453 "spat_L_side" "noBreak"
          movel(spat_L_side_p, a=1.2, v=0.25, r=0.01)
          $ 4454 "spat_L_up" "noBreak"
          movel(spat_L_up_p, a=1.2, v=0.25, r=0.05)
          $ 4455 "MoveJ" "noBreak"
          $ 4456 "Spatula_otw" "noBreak"
          movej(get_inverse_kin(Spatula_otw_p, qnear=Spatula_otw_q), a=1.3962634015954636, v=1.0471975511965976)
        else:
          $ 4457 "ElseIf spatula ≟'spatula_M'" "noBreak"
          if (spatula  == "spatula_M"):
            $ 4458 "MoveJ" "noBreak"
            $ 4459 "Spatula_otw" "noBreak"
            movej(get_inverse_kin(Spatula_otw_p, qnear=Spatula_otw_q), a=1.3962634015954636, v=1.0471975511965976)
            $ 4460 "spat_M_up" "noBreak"
            movej(get_inverse_kin(spat_M_up_p, qnear=spat_M_up_q), a=1.3962634015954636, v=1.0471975511965976, r=0.05)
            $ 4461 "MoveL" "noBreak"
            $ 4462 "spat_M_pick" "noBreak"
            movel(spat_M_pick_p, a=1.2, v=0.25)
            # begin: URCap Program Node
            #   Source: Robotiq_Grippers, 3.17.0.105337, Robotiq Inc.
            #   Type: Gripper
            $ 4463 "Gripper Close (1)" "noBreak"
            if not(gripper_connected[0]):
              popup("Gripper 1 must be connected to run this program.", "No connection", False, True, True)
            end
            if not(rq_is_gripper_activated("1")):
              popup("Gripper 1 is not activated. Go to Installation tab > Gripper to activate it and run the program again.", "Not activated", False, True, True)
            end
            rq_set_pos_spd_for(255, 0, 77, "1")
            rq_wait_pos_spe_for_request(255, 0, 77, "1")
            rq_go_to("1")
            rq_wait("1")
            # end: URCap Program Node
            $ 4464 "spat_M_up" "noBreak"
            movel(spat_M_up_p, a=1.2, v=0.25, r=0.05)
            $ 4465 "Spatula_otw" "noBreak"
            movel(Spatula_otw_p, a=1.2, v=0.25)
            $ 4466 "switch_spat_M≔ False " "noBreak"
            global switch_spat_M=  False
          else:
            $ 4467 "ElseIf spatula≟'spatula_S'" "noBreak"
            if (spatula == "spatula_S"):
              $ 4468 "MoveJ" "noBreak"
              $ 4469 "Spatula_otw" "noBreak"
              movej(get_inverse_kin(Spatula_otw_p, qnear=Spatula_otw_q), a=1.3962634015954636, v=1.0471975511965976)
              $ 4470 "spat_S_Up_7" "noBreak"
              movej(get_inverse_kin(spat_S_Up_7_p, qnear=spat_S_Up_7_q), a=1.3962634015954636, v=1.0471975511965976, r=0.05)
              $ 4471 "MoveL" "noBreak"
              $ 4472 "spat_S_Pick_4" "noBreak"
              movel(spat_S_Pick_4_p, a=1.2, v=0.25)
              # begin: URCap Program Node
              #   Source: Robotiq_Grippers, 3.17.0.105337, Robotiq Inc.
              #   Type: Gripper
              $ 4473 "Gripper Close (1)" "noBreak"
              if not(gripper_connected[0]):
                popup("Gripper 1 must be connected to run this program.", "No connection", False, True, True)
              end
              if not(rq_is_gripper_activated("1")):
                popup("Gripper 1 is not activated. Go to Installation tab > Gripper to activate it and run the program again.", "Not activated", False, True, True)
              end
              rq_set_pos_spd_for(255, 0, 77, "1")
              rq_wait_pos_spe_for_request(255, 0, 77, "1")
              rq_go_to("1")
              rq_wait("1")
              # end: URCap Program Node
              $ 4474 "spat_S_Up_8" "noBreak"
              movel(spat_S_Up_8_p, a=1.2, v=0.25, r=0.05)
              $ 4475 "Spatula_otw" "noBreak"
              movel(Spatula_otw_p, a=1.2, v=0.25)
              $ 4476 "switch_spat_S≔ False " "noBreak"
              global switch_spat_S=  False
            else:
              $ 4477 "ElseIf spatula≟'spatula_flat_M'" "noBreak"
              if (spatula == "spatula_flat_M"):
                $ 4478 "MoveJ" "noBreak"
                $ 4479 "Spatula_otw" "noBreak"
                movej(get_inverse_kin(Spatula_otw_p, qnear=Spatula_otw_q), a=1.3962634015954636, v=1.0471975511965976)
                $ 4480 "spat_flatM_up" "noBreak"
                movej(get_inverse_kin(spat_flatM_up_p, qnear=spat_flatM_up_q), a=1.3962634015954636, v=1.0471975511965976, r=0.05)
                $ 4481 "MoveL" "noBreak"
                $ 4482 "spat_flatM_pick" "noBreak"
                movel(spat_flatM_pick_p, a=1.2, v=0.25)
                # begin: URCap Program Node
                #   Source: Robotiq_Grippers, 3.17.0.105337, Robotiq Inc.
                #   Type: Gripper
                $ 4483 "Gripper Close (1)" "noBreak"
                if not(gripper_connected[0]):
                  popup("Gripper 1 must be connected to run this program.", "No connection", False, True, True)
                end
                if not(rq_is_gripper_activated("1")):
                  popup("Gripper 1 is not activated. Go to Installation tab > Gripper to activate it and run the program again.", "Not activated", False, True, True)
                end
                rq_set_pos_spd_for(255, 0, 77, "1")
                rq_wait_pos_spe_for_request(255, 0, 77, "1")
                rq_go_to("1")
                rq_wait("1")
                # end: URCap Program Node
                $ 4484 "spat_flatM_up" "noBreak"
                movel(spat_flatM_up_p, a=1.2, v=0.25, r=0.05)
                $ 4485 "Spatula_otw" "noBreak"
                movel(Spatula_otw_p, a=1.2, v=0.25)
                $ 4486 "switch_spat_F_M≔ False " "noBreak"
                global switch_spat_F_M=  False
              else:
                $ 4487 "ElseIf spatula≟'spatula_flat_S'" "noBreak"
                if (spatula == "spatula_flat_S"):
                  $ 4488 "MoveJ" "noBreak"
                  $ 4489 "Spatula_otw" "noBreak"
                  movej(get_inverse_kin(Spatula_otw_p, qnear=Spatula_otw_q), a=1.3962634015954636, v=1.0471975511965976)
                  $ 4490 "spat_flatS_up" "noBreak"
                  movej(get_inverse_kin(spat_flatS_up_p, qnear=spat_flatS_up_q), a=1.3962634015954636, v=1.0471975511965976, r=0.05)
                  $ 4491 "MoveL" "noBreak"
                  $ 4492 "spat_flatS_pick" "noBreak"
                  movel(spat_flatS_pick_p, a=1.2, v=0.25)
                  # begin: URCap Program Node
                  #   Source: Robotiq_Grippers, 3.17.0.105337, Robotiq Inc.
                  #   Type: Gripper
                  $ 4493 "Gripper Close (1)" "noBreak"
                  if not(gripper_connected[0]):
                    popup("Gripper 1 must be connected to run this program.", "No connection", False, True, True)
                  end
                  if not(rq_is_gripper_activated("1")):
                    popup("Gripper 1 is not activated. Go to Installation tab > Gripper to activate it and run the program again.", "Not activated", False, True, True)
                  end
                  rq_set_pos_spd_for(255, 0, 77, "1")
                  rq_wait_pos_spe_for_request(255, 0, 77, "1")
                  rq_go_to("1")
                  rq_wait("1")
                  # end: URCap Program Node
                  $ 4494 "spat_flatS_up" "noBreak"
                  movel(spat_flatS_up_p, a=1.2, v=0.25, r=0.05)
                  $ 4495 "Spatula_otw" "noBreak"
                  movel(Spatula_otw_p, a=1.2, v=0.25)
                  $ 4496 "switch_spat_F_S≔ False " "noBreak"
                  global switch_spat_F_S=  False
                end
              end
            end
          end
        end
        $ 4497 "Action_Info≔'Scooping'" "noBreak"
        global Action_Info="Scooping"
        $ 4498 "auto_tilt_and_scoop(W_now, target_weight, weight_value)" "noBreak"
        auto_tilt_and_scoop(W_now, target_weight, weight_value)
        $ 4499 "Action_Info≔'Dosing'" "noBreak"
        global Action_Info="Dosing"
        # begin: URCap Program Node
        #   Source: SensoPart VISOR Robotic, 2.0.6, SensoPart Industriesensorik GmbH
        #   Type: Approach Pose
        $ 4500 "Approach Pose" "noBreak"
        movej(pose_trans(easyPickPose,p[0.0000,0.0000,-0.0000,0.0000,0.0000,0.0000]),a=0.2618,v=0.1745,t=0.000000,r=0.000000)
        # end: URCap Program Node
        # begin: URCap Program Node
        #   Source: SensoPart VISOR Robotic, 2.0.6, SensoPart Industriesensorik GmbH
        #   Type: Target Pose
        $ 4501 "Target Pose" "noBreak"
        movel(pose_trans(easyPickPose,p[0.0000,0.0000,-0.0000,0.0000,0.0000,0.0000]),a=0.0500,v=0.0200,t=0.000000,r=0.000000)
        # end: URCap Program Node
        $ 4502 "Close Gripper" "noBreak"
        $ 4503 "dispense_pos≔get_actual_tcp_pose()" "noBreak"
        global dispense_pos= get_actual_tcp_pose ()
        $ 4504 "Loop weight_value≤target_weight and delta≟0.0 or delta≥0.01" "noBreak"
        thread Thread_while_4504():
          while (True):
            $ 4505 "MoveL" "noBreak"
            $ 4506 "dispense_pos" "noBreak"
            movel(dispense_pos, a=0.2, v=0.1)
            $ 4507 "prev_weight≔get_weight()" "noBreak"
            global prev_weight=get_weight()
            $ 4508 "log_weight()" "noBreak"
            log_weight()
            $ 4509 "Wait: 0.5" "noBreak"
            sleep(0.5)
            $ 4510 "tilt_pose≔pose_trans(get_actual_tcp_pose(), p[0, 0, 0, 0, 0, 2.0])" "noBreak"
            global tilt_pose=pose_trans(get_actual_tcp_pose(), p[0, 0, 0, 0, 0, 2.0])
            $ 4511 "movel(tilt_pose, a=0.5, v=0.5, r=0.00001)" "noBreak"
            movel(tilt_pose, a=0.5, v=0.5, r=0.00001)
            $ 4512 "weight_value≔get_weight()" "noBreak"
            global weight_value=get_weight()
            $ 4513 "tilt_angle≔-1" "noBreak"
            global tilt_angle=-1
            $ 4514 "Wait: 0.5" "noBreak"
            sleep(0.5)
            $ 4515 "dispense_pos" "noBreak"
            movel(dispense_pos, a=1.2, v=0.25)
            $ 4516 "compute_level_percent(W_now, weight_value)" "noBreak"
            compute_level_percent(W_now, weight_value)
            $ 4517 "prev_spat≔spatula" "noBreak"
            global prev_spat=spatula
            $ 4518 "Wait: 0.2" "noBreak"
            sleep(0.2)
            $ 4520 "spatula≔select_spatula(Flowability, level, diff, bulk_density, mouth_d)" "noBreak"
            global spatula=select_spatula(Flowability, level, diff, bulk_density, mouth_d)
            $ 4521 "Wait: 1.0" "noBreak"
            sleep(1.0)
            $ 4522 "send_level_info()" "noBreak"
            send_level_info()
            $ 4523 "send_spatula_info()" "noBreak"
            send_spatula_info()
            $ 4524 "Set AO[0]=0.0" "noBreak"
            set_standard_analog_out(0, 0.0)
            $ 4525 "Wait: 0.5" "noBreak"
            sleep(0.5)
            $ 4526 "swtich spatula" "noBreak"
            $ 4527 "If spatula ≟ 'spatula_M' and switch_spat_M≟ True " "noBreak"
            if (spatula  ==  "spatula_M"  and  switch_spat_M ==   True  ):
              $ 4528 "MoveJ" "noBreak"
              $ 4529 "Spatula_otw" "noBreak"
              movej(get_inverse_kin(Spatula_otw_p, qnear=Spatula_otw_q), a=1.3962634015954636, v=1.0471975511965976)
              $ 4530 "spat_L_up" "noBreak"
              movej(get_inverse_kin(spat_L_up_p, qnear=spat_L_up_q), a=1.3962634015954636, v=1.0471975511965976)
              $ 4531 "MoveL" "noBreak"
              $ 4532 "spat_L_side" "noBreak"
              movel(spat_L_side_p, a=1.2, v=0.25)
              $ 4533 "spat_L_lift" "noBreak"
              movel(spat_L_lift_p, a=1.2, v=0.25)
              $ 4534 "spat_L_pick" "noBreak"
              movel(spat_L_pick_p, a=0.2, v=0.1)
              # begin: URCap Program Node
              #   Source: Robotiq_Grippers, 3.17.0.105337, Robotiq Inc.
              #   Type: Gripper
              $ 4535 "Gripper Open (1)" "noBreak"
              if not(gripper_connected[0]):
                popup("Gripper 1 must be connected to run this program.", "No connection", False, True, True)
              end
              if not(rq_is_gripper_activated("1")):
                popup("Gripper 1 is not activated. Go to Installation tab > Gripper to activate it and run the program again.", "Not activated", False, True, True)
              end
              rq_set_pos_spd_for(0, 255, 77, "1")
              rq_wait_pos_spe_for_request(0, 255, 77, "1")
              rq_go_to("1")
              rq_wait("1")
              # end: URCap Program Node
              $ 4536 "spat_M_pick" "noBreak"
              movel(spat_M_pick_p, a=1.2, v=0.25)
              # begin: URCap Program Node
              #   Source: Robotiq_Grippers, 3.17.0.105337, Robotiq Inc.
              #   Type: Gripper
              $ 4537 "Gripper Close (1)" "noBreak"
              if not(gripper_connected[0]):
                popup("Gripper 1 must be connected to run this program.", "No connection", False, True, True)
              end
              if not(rq_is_gripper_activated("1")):
                popup("Gripper 1 is not activated. Go to Installation tab > Gripper to activate it and run the program again.", "Not activated", False, True, True)
              end
              rq_set_pos_spd_for(255, 0, 77, "1")
              rq_wait_pos_spe_for_request(255, 0, 77, "1")
              rq_go_to("1")
              rq_wait("1")
              # end: URCap Program Node
              $ 4538 "spat_M_up" "noBreak"
              movel(spat_M_up_p, a=1.2, v=0.25)
              $ 4539 "Spatula_otw" "noBreak"
              movel(Spatula_otw_p, a=1.2, v=0.25)
              $ 4540 "switch_spat_M≔ False " "noBreak"
              global switch_spat_M=  False
              $ 4541 "correction_reset()" "noBreak"
              correction_reset()
            else:
              $ 4542 "ElseIf spatula ≟ 'spatula_S' and switch_spat_S ≟ True and prev_spat≟'spatula_M'" "noBreak"
              if (spatula  ==  "spatula_S" and switch_spat_S  ==   True  and prev_spat == "spatula_M"):
                $ 4543 "MoveL" "noBreak"
                $ 4544 "Spatula_otw" "noBreak"
                movel(Spatula_otw_p, a=1.2, v=0.25)
                $ 4545 "spat_M_up" "noBreak"
                movel(spat_M_up_p, a=1.2, v=0.25)
                $ 4546 "spat_M_pick" "noBreak"
                movel(spat_M_pick_p, a=0.2, v=0.1)
                # begin: URCap Program Node
                #   Source: Robotiq_Grippers, 3.17.0.105337, Robotiq Inc.
                #   Type: Gripper
                $ 4547 "Gripper Open (1)" "noBreak"
                if not(gripper_connected[0]):
                  popup("Gripper 1 must be connected to run this program.", "No connection", False, True, True)
                end
                if not(rq_is_gripper_activated("1")):
                  popup("Gripper 1 is not activated. Go to Installation tab > Gripper to activate it and run the program again.", "Not activated", False, True, True)
                end
                rq_set_pos_spd_for(0, 255, 77, "1")
                rq_wait_pos_spe_for_request(0, 255, 77, "1")
                rq_go_to("1")
                rq_wait("1")
                # end: URCap Program Node
                $ 4548 "spat_S_pick" "noBreak"
                movel(spat_S_pick_p, a=1.2, v=0.25)
                # begin: URCap Program Node
                #   Source: Robotiq_Grippers, 3.17.0.105337, Robotiq Inc.
                #   Type: Gripper
                $ 4549 "Gripper Close (1)" "noBreak"
                if not(gripper_connected[0]):
                  popup("Gripper 1 must be connected to run this program.", "No connection", False, True, True)
                end
                if not(rq_is_gripper_activated("1")):
                  popup("Gripper 1 is not activated. Go to Installation tab > Gripper to activate it and run the program again.", "Not activated", False, True, True)
                end
                rq_set_pos_spd_for(255, 0, 77, "1")
                rq_wait_pos_spe_for_request(255, 0, 77, "1")
                rq_go_to("1")
                rq_wait("1")
                # end: URCap Program Node
                $ 4550 "spat_S_up" "noBreak"
                movel(spat_S_up_p, a=1.2, v=0.25)
                $ 4551 "Spatula_otw" "noBreak"
                movel(Spatula_otw_p, a=1.2, v=0.25)
                $ 4552 "switch_spat_S≔ False " "noBreak"
                global switch_spat_S=  False
                $ 4553 "correction_reset()" "noBreak"
                correction_reset()
              else:
                $ 4554 "ElseIf spatula≟'spatula_S' and switch_spat_S≟ True  and prev_spat≟'spatula_L'" "noBreak"
                if (spatula == "spatula_S" and switch_spat_S ==   True    and  prev_spat == "spatula_L"):
                  $ 4555 "MoveJ" "noBreak"
                  $ 4556 "Spatula_otw" "noBreak"
                  movej(get_inverse_kin(Spatula_otw_p, qnear=Spatula_otw_q), a=1.3962634015954636, v=1.0471975511965976)
                  $ 4557 "spat_L_up" "noBreak"
                  movej(get_inverse_kin(spat_L_up_p, qnear=spat_L_up_q), a=1.3962634015954636, v=1.0471975511965976)
                  $ 4558 "MoveL" "noBreak"
                  $ 4559 "spat_L_side" "noBreak"
                  movel(spat_L_side_p, a=1.2, v=0.25)
                  $ 4560 "spat_L_lift" "noBreak"
                  movel(spat_L_lift_p, a=1.2, v=0.25)
                  $ 4561 "spat_L_pick" "noBreak"
                  movel(spat_L_pick_p, a=0.2, v=0.1)
                  # begin: URCap Program Node
                  #   Source: Robotiq_Grippers, 3.17.0.105337, Robotiq Inc.
                  #   Type: Gripper
                  $ 4562 "Gripper Open (1)" "noBreak"
                  if not(gripper_connected[0]):
                    popup("Gripper 1 must be connected to run this program.", "No connection", False, True, True)
                  end
                  if not(rq_is_gripper_activated("1")):
                    popup("Gripper 1 is not activated. Go to Installation tab > Gripper to activate it and run the program again.", "Not activated", False, True, True)
                  end
                  rq_set_pos_spd_for(0, 255, 77, "1")
                  rq_wait_pos_spe_for_request(0, 255, 77, "1")
                  rq_go_to("1")
                  rq_wait("1")
                  # end: URCap Program Node
                  $ 4563 "spat_S_pick" "noBreak"
                  movel(spat_S_pick_p, a=1.2, v=0.25)
                  # begin: URCap Program Node
                  #   Source: Robotiq_Grippers, 3.17.0.105337, Robotiq Inc.
                  #   Type: Gripper
                  $ 4564 "Gripper Close (1)" "noBreak"
                  if not(gripper_connected[0]):
                    popup("Gripper 1 must be connected to run this program.", "No connection", False, True, True)
                  end
                  if not(rq_is_gripper_activated("1")):
                    popup("Gripper 1 is not activated. Go to Installation tab > Gripper to activate it and run the program again.", "Not activated", False, True, True)
                  end
                  rq_set_pos_spd_for(255, 0, 77, "1")
                  rq_wait_pos_spe_for_request(255, 0, 77, "1")
                  rq_go_to("1")
                  rq_wait("1")
                  # end: URCap Program Node
                  $ 4565 "spat_S_up" "noBreak"
                  movel(spat_S_up_p, a=1.2, v=0.25)
                  $ 4566 "Spatula_otw" "noBreak"
                  movel(Spatula_otw_p, a=1.2, v=0.25)
                  $ 4567 "switch_spat_S≔ False " "noBreak"
                  global switch_spat_S=  False
                  $ 4568 "correction_reset()" "noBreak"
                  correction_reset()
                else:
                  $ 4569 "ElseIf spatula≟'spatula_flat_S'  and switch_spat_F_S ≟ True " "noBreak"
                  if (spatula == "spatula_flat_S"   and  switch_spat_F_S  ==   True  ):
                    $ 4570 "MoveL" "noBreak"
                    $ 4571 "Spatula_otw" "noBreak"
                    movel(Spatula_otw_p, a=1.2, v=0.25)
                    $ 4572 "spat_flatM_up" "noBreak"
                    movel(spat_flatM_up_p, a=1.2, v=0.25)
                    $ 4573 "spat_flatM_pick" "noBreak"
                    movel(spat_flatM_pick_p, a=0.2, v=0.1)
                    # begin: URCap Program Node
                    #   Source: Robotiq_Grippers, 3.17.0.105337, Robotiq Inc.
                    #   Type: Gripper
                    $ 4574 "Gripper Open (1)" "noBreak"
                    if not(gripper_connected[0]):
                      popup("Gripper 1 must be connected to run this program.", "No connection", False, True, True)
                    end
                    if not(rq_is_gripper_activated("1")):
                      popup("Gripper 1 is not activated. Go to Installation tab > Gripper to activate it and run the program again.", "Not activated", False, True, True)
                    end
                    rq_set_pos_spd_for(0, 0, 77, "1")
                    rq_wait_pos_spe_for_request(0, 0, 77, "1")
                    rq_go_to("1")
                    rq_wait("1")
                    # end: URCap Program Node
                    $ 4575 "spat_flatS_pick" "noBreak"
                    movel(spat_flatS_pick_p, a=1.2, v=0.25)
                    # begin: URCap Program Node
                    #   Source: Robotiq_Grippers, 3.17.0.105337, Robotiq Inc.
                    #   Type: Gripper
                    $ 4576 "Gripper Close (1)" "noBreak"
                    if not(gripper_connected[0]):
                      popup("Gripper 1 must be connected to run this program.", "No connection", False, True, True)
                    end
                    if not(rq_is_gripper_activated("1")):
                      popup("Gripper 1 is not activated. Go to Installation tab > Gripper to activate it and run the program again.", "Not activated", False, True, True)
                    end
                    rq_set_pos_spd_for(255, 0, 77, "1")
                    rq_wait_pos_spe_for_request(255, 0, 77, "1")
                    rq_go_to("1")
                    rq_wait("1")
                    # end: URCap Program Node
                    $ 4577 "spat_flatS_up" "noBreak"
                    movel(spat_flatS_up_p, a=1.2, v=0.25)
                    $ 4578 "Spatula_otw" "noBreak"
                    movel(Spatula_otw_p, a=1.2, v=0.25)
                    $ 4579 "switch_spat_F_S≔ False " "noBreak"
                    global switch_spat_F_S=  False
                    $ 4580 "correction_reset()" "noBreak"
                    correction_reset()
                  end
                end
              end
            end
            $ 4581 "tilt(level)" "noBreak"
            tilt(level)
            $ 4582 "Action_Info≔'Scooping'" "noBreak"
            global Action_Info="Scooping"
            $ 4583 "auto_tilt_and_scoop(W_now, target_weight, weight_value)" "noBreak"
            auto_tilt_and_scoop(W_now, target_weight, weight_value)
            $ 4584 "Action_Info≔'Dosing'" "noBreak"
            global Action_Info="Dosing"
          end
        end
        if (weight_value <= target_weight and delta == 0.0 or delta >= 0.01):
          global thread_handler_4504=run Thread_while_4504()
